	mF_Mpc_f_a: ARRAY[0..59047] OF LREAL := [-1.7756006070928429E-5, -1.955926027849794E-5, -2.1265642444599059E-5, -2.2878087249309936E-5, -2.4399475238503513E-5, -2.5832632877734329E-5, -2.7180332648224444E-5, -2.8445293182983732E-5, -2.9630179441154765E-5, -3.0737602918726609E-5, -3.1770121893815045E-5, -3.2730241704758869E-5, -3.3620415059333691E-5, -3.4443042373434618E-5, -3.5200472137629193E-5, -3.5895001310030509E-5, -3.652887573398812E-5, -3.7104290579141277E-5, -3.7623390804425058E-5, -3.808827164166491E-5, -3.8500979098439383E-5, -3.886351047893401E-5, -3.9177814921551905E-5, -3.9445793952087749E-5, -3.966930205131298E-5, -3.98501472358593E-5, -3.9990091651326829E-5, -4.0090852176581095E-5, -4.0154101038240283E-5, -4.0181466434390562E-5, -4.017453316660271E-5, -4.013484327935801E-5, -4.0063896706025282E-5, -3.9963151920563813E-5, -3.9834026594159355E-5, -3.9677898256031791E-5, -3.9496104957683613E-5, -3.9289945939888413E-5, -3.9060682301747689E-5, -3.8809537671172525E-5, -3.8537698876174604E-5, -3.8246316616377579E-5, -3.793650613418646E-5, -3.7609347885077623E-5, -3.7265888206497395E-5, -3.6907139984880808E-5, -3.6534083320325723E-5, -3.6147666188480321E-5, -3.5748805099224027E-5, -3.5338385751743129E-5, -3.4917263685623729E-5, -3.44862649276042E-5, -3.40461866336495E-5, -3.3597797726028135E-5, -3.3141839525091535E-5, -3.2679026375472935E-5, -3.221004626644033E-5, -3.1735561446154833E-5, -3.12562090296018E-5, -3.0772601599977736E-5, -3.0285327803331116E-5, -2.9794952936269942E-5, -2.9302019526562752E-5, -2.8807047906473585E-5, -2.8310536778684464E-5, -2.7812963774671571E-5, -2.7314786005413577E-5, -2.6816440604322343E-5, -2.6318345262297408E-5, -2.5820898754816765E-5, -2.5324481460986734E-5, -2.4829455874483883E-5, -2.4336167106331684E-5, -2.3844943379463754E-5, -2.3356096515034559E-5, -2.2869922410446928E-5, -2.2386701509073987E-5, -2.190669926166088E-5, -2.1430166579399207E-5, -2.0957340278674263E-5, -2.0488443517492027E-5, -2.0023686223599328E-5, -1.9563265514316956E-5, -1.910736610811127E-5, -1.8656160727935741E-5, -1.8209810496378919E-5, -1.776846532266075E-5, -1.7332264281523728E-5, -1.6901335984070202E-5, -1.6475798940601218E-5, -1.6055761915516631E-5, -1.5641324274339943E-5, -1.5232576322934952E-5, -1.4829599638984815E-5, -1.4432467395807249E-5, -1.4041244678582621E-5, -1.3655988793074526E-5, -1.3276749566924981E-5, -1.29035696436089E-5, -1.2536484769134677E-5, -1.217552407157984E-5, -1.1820710333552607E-5, -1.1472060257671982E-5, -1.1129584725160594E-5, -1.0793289047645905E-5, -1.0463173212266783E-5, -1.0139232120183559E-5, -9.8214558185907186E-6, -9.5098297263323067E-6, -9.20433485322091E-6, -8.9049480131616991E-6, -8.6116420311836354E-6, -8.324385944480339E-6, -8.04314519756346E-6, -7.7678818316316609E-6, -7.4985546682584246E-6, -7.2351194875019937E-6, -6.9775292005406626E-6, -6.7257340169365817E-6, -6.4796816066309883E-6, 1.7756006070928429E-5, 1.955926027849794E-5, 2.1265642444599059E-5, 2.2878087249309936E-5, 2.4399475238503513E-5, 2.5832632877734329E-5, 2.7180332648224444E-5, 2.8445293182983732E-5, 2.9630179441154765E-5, 3.0737602918726609E-5, 3.1770121893815045E-5, 3.2730241704758869E-5, 3.3620415059333691E-5, 3.4443042373434618E-5, 3.5200472137629193E-5, 3.5895001310030509E-5, 3.652887573398812E-5, 3.7104290579141277E-5, 3.7623390804425058E-5, 3.808827164166491E-5, 3.8500979098439383E-5, 3.886351047893401E-5, 3.9177814921551905E-5, 3.9445793952087749E-5, 3.966930205131298E-5, 3.98501472358593E-5, 3.9990091651326829E-5, 4.0090852176581095E-5, 4.0154101038240283E-5, 4.0181466434390562E-5, 4.017453316660271E-5, 4.013484327935801E-5, 4.0063896706025282E-5, 3.9963151920563813E-5, 3.9834026594159355E-5, 3.9677898256031791E-5, 3.9496104957683613E-5, 3.9289945939888413E-5, 3.9060682301747689E-5, 3.8809537671172525E-5, 3.8537698876174604E-5, 3.8246316616377579E-5, 3.793650613418646E-5, 3.7609347885077623E-5, 3.7265888206497395E-5, 3.6907139984880808E-5, 3.6534083320325723E-5, 3.6147666188480321E-5, 3.5748805099224027E-5, 3.5338385751743129E-5, 3.4917263685623729E-5, 3.44862649276042E-5, 3.40461866336495E-5, 3.3597797726028135E-5, 3.3141839525091535E-5, 3.2679026375472935E-5, 3.221004626644033E-5, 3.1735561446154833E-5, 3.12562090296018E-5, 3.0772601599977736E-5, 3.0285327803331116E-5, 2.9794952936269942E-5, 2.9302019526562752E-5, 2.8807047906473585E-5, 2.8310536778684464E-5, 2.7812963774671571E-5, 2.7314786005413577E-5, 2.6816440604322343E-5, 2.6318345262297408E-5, 2.5820898754816765E-5, 2.5324481460986734E-5, 2.4829455874483883E-5, 2.4336167106331684E-5, 2.3844943379463754E-5, 2.3356096515034559E-5, 2.2869922410446928E-5, 2.2386701509073987E-5, 2.190669926166088E-5, 2.1430166579399207E-5, 2.0957340278674263E-5, 2.0488443517492027E-5, 2.0023686223599328E-5, 1.9563265514316956E-5, 1.910736610811127E-5, 1.8656160727935741E-5, 1.8209810496378919E-5, 1.776846532266075E-5, 1.7332264281523728E-5, 1.6901335984070202E-5, 1.6475798940601218E-5, 1.6055761915516631E-5, 1.5641324274339943E-5, 1.5232576322934952E-5, 1.4829599638984815E-5, 1.4432467395807249E-5, 1.4041244678582621E-5, 1.3655988793074526E-5, 1.3276749566924981E-5, 1.29035696436089E-5, 1.2536484769134677E-5, 1.217552407157984E-5, 1.1820710333552607E-5, 1.1472060257671982E-5, 1.1129584725160594E-5, 1.0793289047645905E-5, 1.0463173212266783E-5, 1.0139232120183559E-5, 9.8214558185907186E-6, 9.5098297263323067E-6, 9.20433485322091E-6, 8.9049480131616991E-6, 8.6116420311836354E-6, 8.324385944480339E-6, 8.04314519756346E-6, 7.7678818316316609E-6, 7.4985546682584246E-6, 7.2351194875019937E-6, 6.9775292005406626E-6, 6.7257340169365817E-6, 6.4796816066309883E-6, 0.0, 0.0, 0.0, 0.0, -0.0, -0.0, -0.0, -0.0, -0.0, -0.0, -0.0, -0.0, -0.0, -0.0, -0.0, -0.0, -0.0, -0.0, -0.0, -0.0, -0.0, -0.0, -0.0, -0.0, -0.0, -0.0, -0.0, -0.0, -0.0, -0.0, -0.0, -0.0, -0.0, -0.0, -0.0, -0.0, -0.0, -0.0, -0.0, -0.0, -0.0, -0.0, -0.0, -0.0, -0.0, -0.0, -0.0, -0.0, -0.0, -0.0, -0.0, -0.0, -0.0, -0.0, -0.0, -0.0, -0.0, -0.0, -0.0, -0.0, -0.0, -0.0, -0.0, -0.0, -0.0, -0.0, -0.0, -0.0, -0.0, -0.0, -0.0, -0.0, -0.0, -0.0, -0.0, -0.0, -0.0, -0.0, -0.0, -0.0, -0.0, -0.0, -0.0, -0.0, -0.0, -0.0, -0.0, -0.0, -0.0, -0.0, -0.0, -0.0, -0.0, -0.0, -0.0, -0.0, -0.0, -0.0, -0.0, -0.0, -0.0, -0.0, -0.0, -0.0, -0.0, -0.0, -0.0, -0.0, -0.0, -0.0, -0.0, -0.0, -0.0, -0.0, -0.0, -0.0, -0.0, -0.0, -0.0, -0.0, -0.0, -0.0, -0.0, -0.0, 0.0, 0.0, 0.0, 0.0, 0.0, 0.0, 0.0, 0.0, 0.0, 0.0, 0.0, 0.0, 0.0, 0.0, 0.0, 0.0, 0.0, 0.0, 0.0, 0.0, 0.0, 0.0, 0.0, 0.0, 0.0, 0.0, 0.0, 0.0, 0.0, 0.0, 0.0, 0.0, 0.0, 0.0, 0.0, 0.0, 0.0, 0.0, 0.0, 0.0, 0.0, 0.0, 0.0, 0.0, 0.0, 0.0, 0.0, 0.0, 0.0, 0.0, 0.0, 0.0, 0.0, 0.0, 0.0, 0.0, 0.0, 0.0, 0.0, 0.0, 0.0, 0.0, 0.0, 0.0, 0.0, 0.0, 0.0, 0.0, 0.0, 0.0, 0.0, 0.0, 0.0, 0.0, 0.0, 0.0, 0.0, 0.0, 0.0, 0.0, 0.0, 0.0, 0.0, 0.0, 0.0, 0.0, 0.0, 0.0, 0.0, 0.0, 0.0, 0.0, 0.0, 0.0, 0.0, 0.0, 0.0, 0.0, 0.0, 0.0, 0.0, 0.0, 0.0, 0.0, 0.0, 0.0, 0.0, 0.0, 0.0, 0.0, 0.0, 0.0, 0.0, 0.0, 0.0, 0.0, 0.0, 0.0, 0.0, 0.0, 0.0, 0.0, 0.0, 0.0, -0.0, -1.7756006070928429E-5, -1.955926027849794E-5, -2.1265642444599059E-5, -2.2878087249309936E-5, -2.4399475238503513E-5, -2.5832632877734329E-5, -2.7180332648224444E-5, -2.8445293182983732E-5, -2.9630179441154765E-5, -3.0737602918726609E-5, -3.1770121893815045E-5, -3.2730241704758869E-5, -3.3620415059333691E-5, -3.4443042373434618E-5, -3.5200472137629193E-5, -3.5895001310030509E-5, -3.652887573398812E-5, -3.7104290579141277E-5, -3.7623390804425058E-5, -3.808827164166491E-5, -3.8500979098439383E-5, -3.886351047893401E-5, -3.9177814921551905E-5, -3.9445793952087749E-5, -3.966930205131298E-5, -3.98501472358593E-5, -3.9990091651326829E-5, -4.0090852176581095E-5, -4.0154101038240283E-5, -4.0181466434390562E-5, -4.017453316660271E-5, -4.013484327935801E-5, -4.0063896706025282E-5, -3.9963151920563813E-5, -3.9834026594159355E-5, -3.9677898256031791E-5, -3.9496104957683613E-5, -3.9289945939888413E-5, -3.9060682301747689E-5, -3.8809537671172525E-5, -3.8537698876174604E-5, -3.8246316616377579E-5, -3.793650613418646E-5, -3.7609347885077623E-5, -3.7265888206497395E-5, -3.6907139984880808E-5, -3.6534083320325723E-5, -3.6147666188480321E-5, -3.5748805099224027E-5, -3.5338385751743129E-5, -3.4917263685623729E-5, -3.44862649276042E-5, -3.40461866336495E-5, -3.3597797726028135E-5, -3.3141839525091535E-5, -3.2679026375472935E-5, -3.221004626644033E-5, -3.1735561446154833E-5, -3.12562090296018E-5, -3.0772601599977736E-5, -3.0285327803331116E-5, -2.9794952936269942E-5, -2.9302019526562752E-5, -2.8807047906473585E-5, -2.8310536778684464E-5, -2.7812963774671571E-5, -2.7314786005413577E-5, -2.6816440604322343E-5, -2.6318345262297408E-5, -2.5820898754816765E-5, -2.5324481460986734E-5, -2.4829455874483883E-5, -2.4336167106331684E-5, -2.3844943379463754E-5, -2.3356096515034559E-5, -2.2869922410446928E-5, -2.2386701509073987E-5, -2.190669926166088E-5, -2.1430166579399207E-5, -2.0957340278674263E-5, -2.0488443517492027E-5, -2.0023686223599328E-5, -1.9563265514316956E-5, -1.910736610811127E-5, -1.8656160727935741E-5, -1.8209810496378919E-5, -1.776846532266075E-5, -1.7332264281523728E-5, -1.6901335984070202E-5, -1.6475798940601218E-5, -1.6055761915516631E-5, -1.5641324274339943E-5, -1.5232576322934952E-5, -1.4829599638984815E-5, -1.4432467395807249E-5, -1.4041244678582621E-5, -1.3655988793074526E-5, -1.3276749566924981E-5, -1.29035696436089E-5, -1.2536484769134677E-5, -1.217552407157984E-5, -1.1820710333552607E-5, -1.1472060257671982E-5, -1.1129584725160594E-5, -1.0793289047645905E-5, -1.0463173212266783E-5, -1.0139232120183559E-5, -9.8214558185907186E-6, -9.5098297263323067E-6, -9.20433485322091E-6, -8.9049480131616991E-6, -8.6116420311836354E-6, -8.324385944480339E-6, -8.04314519756346E-6, -7.7678818316316609E-6, -7.4985546682584246E-6, -7.2351194875019937E-6, -6.9775292005406626E-6, -6.7257340169365817E-6, 0.0, 1.7756006070928429E-5, 1.955926027849794E-5, 2.1265642444599059E-5, 2.2878087249309936E-5, 2.4399475238503513E-5, 2.5832632877734329E-5, 2.7180332648224444E-5, 2.8445293182983732E-5, 2.9630179441154765E-5, 3.0737602918726609E-5, 3.1770121893815045E-5, 3.2730241704758869E-5, 3.3620415059333691E-5, 3.4443042373434618E-5, 3.5200472137629193E-5, 3.5895001310030509E-5, 3.652887573398812E-5, 3.7104290579141277E-5, 3.7623390804425058E-5, 3.808827164166491E-5, 3.8500979098439383E-5, 3.886351047893401E-5, 3.9177814921551905E-5, 3.9445793952087749E-5, 3.966930205131298E-5, 3.98501472358593E-5, 3.9990091651326829E-5, 4.0090852176581095E-5, 4.0154101038240283E-5, 4.0181466434390562E-5, 4.017453316660271E-5, 4.013484327935801E-5, 4.0063896706025282E-5, 3.9963151920563813E-5, 3.9834026594159355E-5, 3.9677898256031791E-5, 3.9496104957683613E-5, 3.9289945939888413E-5, 3.9060682301747689E-5, 3.8809537671172525E-5, 3.8537698876174604E-5, 3.8246316616377579E-5, 3.793650613418646E-5, 3.7609347885077623E-5, 3.7265888206497395E-5, 3.6907139984880808E-5, 3.6534083320325723E-5, 3.6147666188480321E-5, 3.5748805099224027E-5, 3.5338385751743129E-5, 3.4917263685623729E-5, 3.44862649276042E-5, 3.40461866336495E-5, 3.3597797726028135E-5, 3.3141839525091535E-5, 3.2679026375472935E-5, 3.221004626644033E-5, 3.1735561446154833E-5, 3.12562090296018E-5, 3.0772601599977736E-5, 3.0285327803331116E-5, 2.9794952936269942E-5, 2.9302019526562752E-5, 2.8807047906473585E-5, 2.8310536778684464E-5, 2.7812963774671571E-5, 2.7314786005413577E-5, 2.6816440604322343E-5, 2.6318345262297408E-5, 2.5820898754816765E-5, 2.5324481460986734E-5, 2.4829455874483883E-5, 2.4336167106331684E-5, 2.3844943379463754E-5, 2.3356096515034559E-5, 2.2869922410446928E-5, 2.2386701509073987E-5, 2.190669926166088E-5, 2.1430166579399207E-5, 2.0957340278674263E-5, 2.0488443517492027E-5, 2.0023686223599328E-5, 1.9563265514316956E-5, 1.910736610811127E-5, 1.8656160727935741E-5, 1.8209810496378919E-5, 1.776846532266075E-5, 1.7332264281523728E-5, 1.6901335984070202E-5, 1.6475798940601218E-5, 1.6055761915516631E-5, 1.5641324274339943E-5, 1.5232576322934952E-5, 1.4829599638984815E-5, 1.4432467395807249E-5, 1.4041244678582621E-5, 1.3655988793074526E-5, 1.3276749566924981E-5, 1.29035696436089E-5, 1.2536484769134677E-5, 1.217552407157984E-5, 1.1820710333552607E-5, 1.1472060257671982E-5, 1.1129584725160594E-5, 1.0793289047645905E-5, 1.0463173212266783E-5, 1.0139232120183559E-5, 9.8214558185907186E-6, 9.5098297263323067E-6, 9.20433485322091E-6, 8.9049480131616991E-6, 8.6116420311836354E-6, 8.324385944480339E-6, 8.04314519756346E-6, 7.7678818316316609E-6, 7.4985546682584246E-6, 7.2351194875019937E-6, 6.9775292005406626E-6, 6.7257340169365817E-6, 0.0, 0.0, 0.0, 0.0, -0.0, -0.0, -0.0, -0.0, -0.0, -0.0, -0.0, -0.0, -0.0, -0.0, -0.0, -0.0, -0.0, -0.0, -0.0, -0.0, -0.0, -0.0, -0.0, -0.0, -0.0, -0.0, -0.0, -0.0, -0.0, -0.0, -0.0, -0.0, -0.0, -0.0, -0.0, -0.0, -0.0, -0.0, -0.0, -0.0, -0.0, -0.0, -0.0, -0.0, -0.0, -0.0, -0.0, -0.0, -0.0, -0.0, -0.0, -0.0, -0.0, -0.0, -0.0, -0.0, -0.0, -0.0, -0.0, -0.0, -0.0, -0.0, -0.0, -0.0, -0.0, -0.0, -0.0, -0.0, -0.0, -0.0, -0.0, -0.0, -0.0, -0.0, -0.0, -0.0, -0.0, -0.0, -0.0, -0.0, -0.0, -0.0, -0.0, -0.0, -0.0, -0.0, -0.0, -0.0, -0.0, -0.0, -0.0, -0.0, -0.0, -0.0, -0.0, -0.0, -0.0, -0.0, -0.0, -0.0, -0.0, -0.0, -0.0, -0.0, -0.0, -0.0, -0.0, -0.0, -0.0, -0.0, -0.0, -0.0, -0.0, -0.0, -0.0, -0.0, -0.0, -0.0, -0.0, -0.0, -0.0, -0.0, -0.0, -0.0, 0.0, 0.0, 0.0, 0.0, 0.0, 0.0, 0.0, 0.0, 0.0, 0.0, 0.0, 0.0, 0.0, 0.0, 0.0, 0.0, 0.0, 0.0, 0.0, 0.0, 0.0, 0.0, 0.0, 0.0, 0.0, 0.0, 0.0, 0.0, 0.0, 0.0, 0.0, 0.0, 0.0, 0.0, 0.0, 0.0, 0.0, 0.0, 0.0, 0.0, 0.0, 0.0, 0.0, 0.0, 0.0, 0.0, 0.0, 0.0, 0.0, 0.0, 0.0, 0.0, 0.0, 0.0, 0.0, 0.0, 0.0, 0.0, 0.0, 0.0, 0.0, 0.0, 0.0, 0.0, 0.0, 0.0, 0.0, 0.0, 0.0, 0.0, 0.0, 0.0, 0.0, 0.0, 0.0, 0.0, 0.0, 0.0, 0.0, 0.0, 0.0, 0.0, 0.0, 0.0, 0.0, 0.0, 0.0, 0.0, 0.0, 0.0, 0.0, 0.0, 0.0, 0.0, 0.0, 0.0, 0.0, 0.0, 0.0, 0.0, 0.0, 0.0, 0.0, 0.0, 0.0, 0.0, 0.0, 0.0, 0.0, 0.0, 0.0, 0.0, 0.0, 0.0, 0.0, 0.0, 0.0, 0.0, 0.0, 0.0, 0.0, 0.0, 0.0, 0.0, -0.0, -0.0, -1.7756006070928429E-5, -1.955926027849794E-5, -2.1265642444599059E-5, -2.2878087249309936E-5, -2.4399475238503513E-5, -2.5832632877734329E-5, -2.7180332648224444E-5, -2.8445293182983732E-5, -2.9630179441154765E-5, -3.0737602918726609E-5, -3.1770121893815045E-5, -3.2730241704758869E-5, -3.3620415059333691E-5, -3.4443042373434618E-5, -3.5200472137629193E-5, -3.5895001310030509E-5, -3.652887573398812E-5, -3.7104290579141277E-5, -3.7623390804425058E-5, -3.808827164166491E-5, -3.8500979098439383E-5, -3.886351047893401E-5, -3.9177814921551905E-5, -3.9445793952087749E-5, -3.966930205131298E-5, -3.98501472358593E-5, -3.9990091651326829E-5, -4.0090852176581095E-5, -4.0154101038240283E-5, -4.0181466434390562E-5, -4.017453316660271E-5, -4.013484327935801E-5, -4.0063896706025282E-5, -3.9963151920563813E-5, -3.9834026594159355E-5, -3.9677898256031791E-5, -3.9496104957683613E-5, -3.9289945939888413E-5, -3.9060682301747689E-5, -3.8809537671172525E-5, -3.8537698876174604E-5, -3.8246316616377579E-5, -3.793650613418646E-5, -3.7609347885077623E-5, -3.7265888206497395E-5, -3.6907139984880808E-5, -3.6534083320325723E-5, -3.6147666188480321E-5, -3.5748805099224027E-5, -3.5338385751743129E-5, -3.4917263685623729E-5, -3.44862649276042E-5, -3.40461866336495E-5, -3.3597797726028135E-5, -3.3141839525091535E-5, -3.2679026375472935E-5, -3.221004626644033E-5, -3.1735561446154833E-5, -3.12562090296018E-5, -3.0772601599977736E-5, -3.0285327803331116E-5, -2.9794952936269942E-5, -2.9302019526562752E-5, -2.8807047906473585E-5, -2.8310536778684464E-5, -2.7812963774671571E-5, -2.7314786005413577E-5, -2.6816440604322343E-5, -2.6318345262297408E-5, -2.5820898754816765E-5, -2.5324481460986734E-5, -2.4829455874483883E-5, -2.4336167106331684E-5, -2.3844943379463754E-5, -2.3356096515034559E-5, -2.2869922410446928E-5, -2.2386701509073987E-5, -2.190669926166088E-5, -2.1430166579399207E-5, -2.0957340278674263E-5, -2.0488443517492027E-5, -2.0023686223599328E-5, -1.9563265514316956E-5, -1.910736610811127E-5, -1.8656160727935741E-5, -1.8209810496378919E-5, -1.776846532266075E-5, -1.7332264281523728E-5, -1.6901335984070202E-5, -1.6475798940601218E-5, -1.6055761915516631E-5, -1.5641324274339943E-5, -1.5232576322934952E-5, -1.4829599638984815E-5, -1.4432467395807249E-5, -1.4041244678582621E-5, -1.3655988793074526E-5, -1.3276749566924981E-5, -1.29035696436089E-5, -1.2536484769134677E-5, -1.217552407157984E-5, -1.1820710333552607E-5, -1.1472060257671982E-5, -1.1129584725160594E-5, -1.0793289047645905E-5, -1.0463173212266783E-5, -1.0139232120183559E-5, -9.8214558185907186E-6, -9.5098297263323067E-6, -9.20433485322091E-6, -8.9049480131616991E-6, -8.6116420311836354E-6, -8.324385944480339E-6, -8.04314519756346E-6, -7.7678818316316609E-6, -7.4985546682584246E-6, -7.2351194875019937E-6, -6.9775292005406626E-6, 0.0, 0.0, 1.7756006070928429E-5, 1.955926027849794E-5, 2.1265642444599059E-5, 2.2878087249309936E-5, 2.4399475238503513E-5, 2.5832632877734329E-5, 2.7180332648224444E-5, 2.8445293182983732E-5, 2.9630179441154765E-5, 3.0737602918726609E-5, 3.1770121893815045E-5, 3.2730241704758869E-5, 3.3620415059333691E-5, 3.4443042373434618E-5, 3.5200472137629193E-5, 3.5895001310030509E-5, 3.652887573398812E-5, 3.7104290579141277E-5, 3.7623390804425058E-5, 3.808827164166491E-5, 3.8500979098439383E-5, 3.886351047893401E-5, 3.9177814921551905E-5, 3.9445793952087749E-5, 3.966930205131298E-5, 3.98501472358593E-5, 3.9990091651326829E-5, 4.0090852176581095E-5, 4.0154101038240283E-5, 4.0181466434390562E-5, 4.017453316660271E-5, 4.013484327935801E-5, 4.0063896706025282E-5, 3.9963151920563813E-5, 3.9834026594159355E-5, 3.9677898256031791E-5, 3.9496104957683613E-5, 3.9289945939888413E-5, 3.9060682301747689E-5, 3.8809537671172525E-5, 3.8537698876174604E-5, 3.8246316616377579E-5, 3.793650613418646E-5, 3.7609347885077623E-5, 3.7265888206497395E-5, 3.6907139984880808E-5, 3.6534083320325723E-5, 3.6147666188480321E-5, 3.5748805099224027E-5, 3.5338385751743129E-5, 3.4917263685623729E-5, 3.44862649276042E-5, 3.40461866336495E-5, 3.3597797726028135E-5, 3.3141839525091535E-5, 3.2679026375472935E-5, 3.221004626644033E-5, 3.1735561446154833E-5, 3.12562090296018E-5, 3.0772601599977736E-5, 3.0285327803331116E-5, 2.9794952936269942E-5, 2.9302019526562752E-5, 2.8807047906473585E-5, 2.8310536778684464E-5, 2.7812963774671571E-5, 2.7314786005413577E-5, 2.6816440604322343E-5, 2.6318345262297408E-5, 2.5820898754816765E-5, 2.5324481460986734E-5, 2.4829455874483883E-5, 2.4336167106331684E-5, 2.3844943379463754E-5, 2.3356096515034559E-5, 2.2869922410446928E-5, 2.2386701509073987E-5, 2.190669926166088E-5, 2.1430166579399207E-5, 2.0957340278674263E-5, 2.0488443517492027E-5, 2.0023686223599328E-5, 1.9563265514316956E-5, 1.910736610811127E-5, 1.8656160727935741E-5, 1.8209810496378919E-5, 1.776846532266075E-5, 1.7332264281523728E-5, 1.6901335984070202E-5, 1.6475798940601218E-5, 1.6055761915516631E-5, 1.5641324274339943E-5, 1.5232576322934952E-5, 1.4829599638984815E-5, 1.4432467395807249E-5, 1.4041244678582621E-5, 1.3655988793074526E-5, 1.3276749566924981E-5, 1.29035696436089E-5, 1.2536484769134677E-5, 1.217552407157984E-5, 1.1820710333552607E-5, 1.1472060257671982E-5, 1.1129584725160594E-5, 1.0793289047645905E-5, 1.0463173212266783E-5, 1.0139232120183559E-5, 9.8214558185907186E-6, 9.5098297263323067E-6, 9.20433485322091E-6, 8.9049480131616991E-6, 8.6116420311836354E-6, 8.324385944480339E-6, 8.04314519756346E-6, 7.7678818316316609E-6, 7.4985546682584246E-6, 7.2351194875019937E-6, 6.9775292005406626E-6, 0.0, 0.0, 0.0, 0.0, -0.0, -0.0, -0.0, -0.0, -0.0, -0.0, -0.0, -0.0, -0.0, -0.0, -0.0, -0.0, -0.0, -0.0, -0.0, -0.0, -0.0, -0.0, -0.0, -0.0, -0.0, -0.0, -0.0, -0.0, -0.0, -0.0, -0.0, -0.0, -0.0, -0.0, -0.0, -0.0, -0.0, -0.0, -0.0, -0.0, -0.0, -0.0, -0.0, -0.0, -0.0, -0.0, -0.0, -0.0, -0.0, -0.0, -0.0, -0.0, -0.0, -0.0, -0.0, -0.0, -0.0, -0.0, -0.0, -0.0, -0.0, -0.0, -0.0, -0.0, -0.0, -0.0, -0.0, -0.0, -0.0, -0.0, -0.0, -0.0, -0.0, -0.0, -0.0, -0.0, -0.0, -0.0, -0.0, -0.0, -0.0, -0.0, -0.0, -0.0, -0.0, -0.0, -0.0, -0.0, -0.0, -0.0, -0.0, -0.0, -0.0, -0.0, -0.0, -0.0, -0.0, -0.0, -0.0, -0.0, -0.0, -0.0, -0.0, -0.0, -0.0, -0.0, -0.0, -0.0, -0.0, -0.0, -0.0, -0.0, -0.0, -0.0, -0.0, -0.0, -0.0, -0.0, -0.0, -0.0, -0.0, -0.0, -0.0, -0.0, 0.0, 0.0, 0.0, 0.0, 0.0, 0.0, 0.0, 0.0, 0.0, 0.0, 0.0, 0.0, 0.0, 0.0, 0.0, 0.0, 0.0, 0.0, 0.0, 0.0, 0.0, 0.0, 0.0, 0.0, 0.0, 0.0, 0.0, 0.0, 0.0, 0.0, 0.0, 0.0, 0.0, 0.0, 0.0, 0.0, 0.0, 0.0, 0.0, 0.0, 0.0, 0.0, 0.0, 0.0, 0.0, 0.0, 0.0, 0.0, 0.0, 0.0, 0.0, 0.0, 0.0, 0.0, 0.0, 0.0, 0.0, 0.0, 0.0, 0.0, 0.0, 0.0, 0.0, 0.0, 0.0, 0.0, 0.0, 0.0, 0.0, 0.0, 0.0, 0.0, 0.0, 0.0, 0.0, 0.0, 0.0, 0.0, 0.0, 0.0, 0.0, 0.0, 0.0, 0.0, 0.0, 0.0, 0.0, 0.0, 0.0, 0.0, 0.0, 0.0, 0.0, 0.0, 0.0, 0.0, 0.0, 0.0, 0.0, 0.0, 0.0, 0.0, 0.0, 0.0, 0.0, 0.0, 0.0, 0.0, 0.0, 0.0, 0.0, 0.0, 0.0, 0.0, 0.0, 0.0, 0.0, 0.0, 0.0, 0.0, 0.0, 0.0, 0.0, 0.0, -0.0, -0.0, -0.0, -1.7756006070928429E-5, -1.955926027849794E-5, -2.1265642444599059E-5, -2.2878087249309936E-5, -2.4399475238503513E-5, -2.5832632877734329E-5, -2.7180332648224444E-5, -2.8445293182983732E-5, -2.9630179441154765E-5, -3.0737602918726609E-5, -3.1770121893815045E-5, -3.2730241704758869E-5, -3.3620415059333691E-5, -3.4443042373434618E-5, -3.5200472137629193E-5, -3.5895001310030509E-5, -3.652887573398812E-5, -3.7104290579141277E-5, -3.7623390804425058E-5, -3.808827164166491E-5, -3.8500979098439383E-5, -3.886351047893401E-5, -3.9177814921551905E-5, -3.9445793952087749E-5, -3.966930205131298E-5, -3.98501472358593E-5, -3.9990091651326829E-5, -4.0090852176581095E-5, -4.0154101038240283E-5, -4.0181466434390562E-5, -4.017453316660271E-5, -4.013484327935801E-5, -4.0063896706025282E-5, -3.9963151920563813E-5, -3.9834026594159355E-5, -3.9677898256031791E-5, -3.9496104957683613E-5, -3.9289945939888413E-5, -3.9060682301747689E-5, -3.8809537671172525E-5, -3.8537698876174604E-5, -3.8246316616377579E-5, -3.793650613418646E-5, -3.7609347885077623E-5, -3.7265888206497395E-5, -3.6907139984880808E-5, -3.6534083320325723E-5, -3.6147666188480321E-5, -3.5748805099224027E-5, -3.5338385751743129E-5, -3.4917263685623729E-5, -3.44862649276042E-5, -3.40461866336495E-5, -3.3597797726028135E-5, -3.3141839525091535E-5, -3.2679026375472935E-5, -3.221004626644033E-5, -3.1735561446154833E-5, -3.12562090296018E-5, -3.0772601599977736E-5, -3.0285327803331116E-5, -2.9794952936269942E-5, -2.9302019526562752E-5, -2.8807047906473585E-5, -2.8310536778684464E-5, -2.7812963774671571E-5, -2.7314786005413577E-5, -2.6816440604322343E-5, -2.6318345262297408E-5, -2.5820898754816765E-5, -2.5324481460986734E-5, -2.4829455874483883E-5, -2.4336167106331684E-5, -2.3844943379463754E-5, -2.3356096515034559E-5, -2.2869922410446928E-5, -2.2386701509073987E-5, -2.190669926166088E-5, -2.1430166579399207E-5, -2.0957340278674263E-5, -2.0488443517492027E-5, -2.0023686223599328E-5, -1.9563265514316956E-5, -1.910736610811127E-5, -1.8656160727935741E-5, -1.8209810496378919E-5, -1.776846532266075E-5, -1.7332264281523728E-5, -1.6901335984070202E-5, -1.6475798940601218E-5, -1.6055761915516631E-5, -1.5641324274339943E-5, -1.5232576322934952E-5, -1.4829599638984815E-5, -1.4432467395807249E-5, -1.4041244678582621E-5, -1.3655988793074526E-5, -1.3276749566924981E-5, -1.29035696436089E-5, -1.2536484769134677E-5, -1.217552407157984E-5, -1.1820710333552607E-5, -1.1472060257671982E-5, -1.1129584725160594E-5, -1.0793289047645905E-5, -1.0463173212266783E-5, -1.0139232120183559E-5, -9.8214558185907186E-6, -9.5098297263323067E-6, -9.20433485322091E-6, -8.9049480131616991E-6, -8.6116420311836354E-6, -8.324385944480339E-6, -8.04314519756346E-6, -7.7678818316316609E-6, -7.4985546682584246E-6, -7.2351194875019937E-6, 0.0, 0.0, 0.0, 1.7756006070928429E-5, 1.955926027849794E-5, 2.1265642444599059E-5, 2.2878087249309936E-5, 2.4399475238503513E-5, 2.5832632877734329E-5, 2.7180332648224444E-5, 2.8445293182983732E-5, 2.9630179441154765E-5, 3.0737602918726609E-5, 3.1770121893815045E-5, 3.2730241704758869E-5, 3.3620415059333691E-5, 3.4443042373434618E-5, 3.5200472137629193E-5, 3.5895001310030509E-5, 3.652887573398812E-5, 3.7104290579141277E-5, 3.7623390804425058E-5, 3.808827164166491E-5, 3.8500979098439383E-5, 3.886351047893401E-5, 3.9177814921551905E-5, 3.9445793952087749E-5, 3.966930205131298E-5, 3.98501472358593E-5, 3.9990091651326829E-5, 4.0090852176581095E-5, 4.0154101038240283E-5, 4.0181466434390562E-5, 4.017453316660271E-5, 4.013484327935801E-5, 4.0063896706025282E-5, 3.9963151920563813E-5, 3.9834026594159355E-5, 3.9677898256031791E-5, 3.9496104957683613E-5, 3.9289945939888413E-5, 3.9060682301747689E-5, 3.8809537671172525E-5, 3.8537698876174604E-5, 3.8246316616377579E-5, 3.793650613418646E-5, 3.7609347885077623E-5, 3.7265888206497395E-5, 3.6907139984880808E-5, 3.6534083320325723E-5, 3.6147666188480321E-5, 3.5748805099224027E-5, 3.5338385751743129E-5, 3.4917263685623729E-5, 3.44862649276042E-5, 3.40461866336495E-5, 3.3597797726028135E-5, 3.3141839525091535E-5, 3.2679026375472935E-5, 3.221004626644033E-5, 3.1735561446154833E-5, 3.12562090296018E-5, 3.0772601599977736E-5, 3.0285327803331116E-5, 2.9794952936269942E-5, 2.9302019526562752E-5, 2.8807047906473585E-5, 2.8310536778684464E-5, 2.7812963774671571E-5, 2.7314786005413577E-5, 2.6816440604322343E-5, 2.6318345262297408E-5, 2.5820898754816765E-5, 2.5324481460986734E-5, 2.4829455874483883E-5, 2.4336167106331684E-5, 2.3844943379463754E-5, 2.3356096515034559E-5, 2.2869922410446928E-5, 2.2386701509073987E-5, 2.190669926166088E-5, 2.1430166579399207E-5, 2.0957340278674263E-5, 2.0488443517492027E-5, 2.0023686223599328E-5, 1.9563265514316956E-5, 1.910736610811127E-5, 1.8656160727935741E-5, 1.8209810496378919E-5, 1.776846532266075E-5, 1.7332264281523728E-5, 1.6901335984070202E-5, 1.6475798940601218E-5, 1.6055761915516631E-5, 1.5641324274339943E-5, 1.5232576322934952E-5, 1.4829599638984815E-5, 1.4432467395807249E-5, 1.4041244678582621E-5, 1.3655988793074526E-5, 1.3276749566924981E-5, 1.29035696436089E-5, 1.2536484769134677E-5, 1.217552407157984E-5, 1.1820710333552607E-5, 1.1472060257671982E-5, 1.1129584725160594E-5, 1.0793289047645905E-5, 1.0463173212266783E-5, 1.0139232120183559E-5, 9.8214558185907186E-6, 9.5098297263323067E-6, 9.20433485322091E-6, 8.9049480131616991E-6, 8.6116420311836354E-6, 8.324385944480339E-6, 8.04314519756346E-6, 7.7678818316316609E-6, 7.4985546682584246E-6, 7.2351194875019937E-6, 0.0, 0.0, 0.0, 0.0, -0.0, -0.0, -0.0, -0.0, -0.0, -0.0, -0.0, -0.0, -0.0, -0.0, -0.0, -0.0, -0.0, -0.0, -0.0, -0.0, -0.0, -0.0, -0.0, -0.0, -0.0, -0.0, -0.0, -0.0, -0.0, -0.0, -0.0, -0.0, -0.0, -0.0, -0.0, -0.0, -0.0, -0.0, -0.0, -0.0, -0.0, -0.0, -0.0, -0.0, -0.0, -0.0, -0.0, -0.0, -0.0, -0.0, -0.0, -0.0, -0.0, -0.0, -0.0, -0.0, -0.0, -0.0, -0.0, -0.0, -0.0, -0.0, -0.0, -0.0, -0.0, -0.0, -0.0, -0.0, -0.0, -0.0, -0.0, -0.0, -0.0, -0.0, -0.0, -0.0, -0.0, -0.0, -0.0, -0.0, -0.0, -0.0, -0.0, -0.0, -0.0, -0.0, -0.0, -0.0, -0.0, -0.0, -0.0, -0.0, -0.0, -0.0, -0.0, -0.0, -0.0, -0.0, -0.0, -0.0, -0.0, -0.0, -0.0, -0.0, -0.0, -0.0, -0.0, -0.0, -0.0, -0.0, -0.0, -0.0, -0.0, -0.0, -0.0, -0.0, -0.0, -0.0, -0.0, -0.0, -0.0, -0.0, -0.0, -0.0, 0.0, 0.0, 0.0, 0.0, 0.0, 0.0, 0.0, 0.0, 0.0, 0.0, 0.0, 0.0, 0.0, 0.0, 0.0, 0.0, 0.0, 0.0, 0.0, 0.0, 0.0, 0.0, 0.0, 0.0, 0.0, 0.0, 0.0, 0.0, 0.0, 0.0, 0.0, 0.0, 0.0, 0.0, 0.0, 0.0, 0.0, 0.0, 0.0, 0.0, 0.0, 0.0, 0.0, 0.0, 0.0, 0.0, 0.0, 0.0, 0.0, 0.0, 0.0, 0.0, 0.0, 0.0, 0.0, 0.0, 0.0, 0.0, 0.0, 0.0, 0.0, 0.0, 0.0, 0.0, 0.0, 0.0, 0.0, 0.0, 0.0, 0.0, 0.0, 0.0, 0.0, 0.0, 0.0, 0.0, 0.0, 0.0, 0.0, 0.0, 0.0, 0.0, 0.0, 0.0, 0.0, 0.0, 0.0, 0.0, 0.0, 0.0, 0.0, 0.0, 0.0, 0.0, 0.0, 0.0, 0.0, 0.0, 0.0, 0.0, 0.0, 0.0, 0.0, 0.0, 0.0, 0.0, 0.0, 0.0, 0.0, 0.0, 0.0, 0.0, 0.0, 0.0, 0.0, 0.0, 0.0, 0.0, 0.0, 0.0, 0.0, 0.0, 0.0, 0.0, -0.0, -0.0, -0.0, -0.0, -1.7756006070928429E-5, -1.955926027849794E-5, -2.1265642444599059E-5, -2.2878087249309936E-5, -2.4399475238503513E-5, -2.5832632877734329E-5, -2.7180332648224444E-5, -2.8445293182983732E-5, -2.9630179441154765E-5, -3.0737602918726609E-5, -3.1770121893815045E-5, -3.2730241704758869E-5, -3.3620415059333691E-5, -3.4443042373434618E-5, -3.5200472137629193E-5, -3.5895001310030509E-5, -3.652887573398812E-5, -3.7104290579141277E-5, -3.7623390804425058E-5, -3.808827164166491E-5, -3.8500979098439383E-5, -3.886351047893401E-5, -3.9177814921551905E-5, -3.9445793952087749E-5, -3.966930205131298E-5, -3.98501472358593E-5, -3.9990091651326829E-5, -4.0090852176581095E-5, -4.0154101038240283E-5, -4.0181466434390562E-5, -4.017453316660271E-5, -4.013484327935801E-5, -4.0063896706025282E-5, -3.9963151920563813E-5, -3.9834026594159355E-5, -3.9677898256031791E-5, -3.9496104957683613E-5, -3.9289945939888413E-5, -3.9060682301747689E-5, -3.8809537671172525E-5, -3.8537698876174604E-5, -3.8246316616377579E-5, -3.793650613418646E-5, -3.7609347885077623E-5, -3.7265888206497395E-5, -3.6907139984880808E-5, -3.6534083320325723E-5, -3.6147666188480321E-5, -3.5748805099224027E-5, -3.5338385751743129E-5, -3.4917263685623729E-5, -3.44862649276042E-5, -3.40461866336495E-5, -3.3597797726028135E-5, -3.3141839525091535E-5, -3.2679026375472935E-5, -3.221004626644033E-5, -3.1735561446154833E-5, -3.12562090296018E-5, -3.0772601599977736E-5, -3.0285327803331116E-5, -2.9794952936269942E-5, -2.9302019526562752E-5, -2.8807047906473585E-5, -2.8310536778684464E-5, -2.7812963774671571E-5, -2.7314786005413577E-5, -2.6816440604322343E-5, -2.6318345262297408E-5, -2.5820898754816765E-5, -2.5324481460986734E-5, -2.4829455874483883E-5, -2.4336167106331684E-5, -2.3844943379463754E-5, -2.3356096515034559E-5, -2.2869922410446928E-5, -2.2386701509073987E-5, -2.190669926166088E-5, -2.1430166579399207E-5, -2.0957340278674263E-5, -2.0488443517492027E-5, -2.0023686223599328E-5, -1.9563265514316956E-5, -1.910736610811127E-5, -1.8656160727935741E-5, -1.8209810496378919E-5, -1.776846532266075E-5, -1.7332264281523728E-5, -1.6901335984070202E-5, -1.6475798940601218E-5, -1.6055761915516631E-5, -1.5641324274339943E-5, -1.5232576322934952E-5, -1.4829599638984815E-5, -1.4432467395807249E-5, -1.4041244678582621E-5, -1.3655988793074526E-5, -1.3276749566924981E-5, -1.29035696436089E-5, -1.2536484769134677E-5, -1.217552407157984E-5, -1.1820710333552607E-5, -1.1472060257671982E-5, -1.1129584725160594E-5, -1.0793289047645905E-5, -1.0463173212266783E-5, -1.0139232120183559E-5, -9.8214558185907186E-6, -9.5098297263323067E-6, -9.20433485322091E-6, -8.9049480131616991E-6, -8.6116420311836354E-6, -8.324385944480339E-6, -8.04314519756346E-6, -7.7678818316316609E-6, -7.4985546682584246E-6, 0.0, 0.0, 0.0, 0.0, 1.7756006070928429E-5, 1.955926027849794E-5, 2.1265642444599059E-5, 2.2878087249309936E-5, 2.4399475238503513E-5, 2.5832632877734329E-5, 2.7180332648224444E-5, 2.8445293182983732E-5, 2.9630179441154765E-5, 3.0737602918726609E-5, 3.1770121893815045E-5, 3.2730241704758869E-5, 3.3620415059333691E-5, 3.4443042373434618E-5, 3.5200472137629193E-5, 3.5895001310030509E-5, 3.652887573398812E-5, 3.7104290579141277E-5, 3.7623390804425058E-5, 3.808827164166491E-5, 3.8500979098439383E-5, 3.886351047893401E-5, 3.9177814921551905E-5, 3.9445793952087749E-5, 3.966930205131298E-5, 3.98501472358593E-5, 3.9990091651326829E-5, 4.0090852176581095E-5, 4.0154101038240283E-5, 4.0181466434390562E-5, 4.017453316660271E-5, 4.013484327935801E-5, 4.0063896706025282E-5, 3.9963151920563813E-5, 3.9834026594159355E-5, 3.9677898256031791E-5, 3.9496104957683613E-5, 3.9289945939888413E-5, 3.9060682301747689E-5, 3.8809537671172525E-5, 3.8537698876174604E-5, 3.8246316616377579E-5, 3.793650613418646E-5, 3.7609347885077623E-5, 3.7265888206497395E-5, 3.6907139984880808E-5, 3.6534083320325723E-5, 3.6147666188480321E-5, 3.5748805099224027E-5, 3.5338385751743129E-5, 3.4917263685623729E-5, 3.44862649276042E-5, 3.40461866336495E-5, 3.3597797726028135E-5, 3.3141839525091535E-5, 3.2679026375472935E-5, 3.221004626644033E-5, 3.1735561446154833E-5, 3.12562090296018E-5, 3.0772601599977736E-5, 3.0285327803331116E-5, 2.9794952936269942E-5, 2.9302019526562752E-5, 2.8807047906473585E-5, 2.8310536778684464E-5, 2.7812963774671571E-5, 2.7314786005413577E-5, 2.6816440604322343E-5, 2.6318345262297408E-5, 2.5820898754816765E-5, 2.5324481460986734E-5, 2.4829455874483883E-5, 2.4336167106331684E-5, 2.3844943379463754E-5, 2.3356096515034559E-5, 2.2869922410446928E-5, 2.2386701509073987E-5, 2.190669926166088E-5, 2.1430166579399207E-5, 2.0957340278674263E-5, 2.0488443517492027E-5, 2.0023686223599328E-5, 1.9563265514316956E-5, 1.910736610811127E-5, 1.8656160727935741E-5, 1.8209810496378919E-5, 1.776846532266075E-5, 1.7332264281523728E-5, 1.6901335984070202E-5, 1.6475798940601218E-5, 1.6055761915516631E-5, 1.5641324274339943E-5, 1.5232576322934952E-5, 1.4829599638984815E-5, 1.4432467395807249E-5, 1.4041244678582621E-5, 1.3655988793074526E-5, 1.3276749566924981E-5, 1.29035696436089E-5, 1.2536484769134677E-5, 1.217552407157984E-5, 1.1820710333552607E-5, 1.1472060257671982E-5, 1.1129584725160594E-5, 1.0793289047645905E-5, 1.0463173212266783E-5, 1.0139232120183559E-5, 9.8214558185907186E-6, 9.5098297263323067E-6, 9.20433485322091E-6, 8.9049480131616991E-6, 8.6116420311836354E-6, 8.324385944480339E-6, 8.04314519756346E-6, 7.7678818316316609E-6, 7.4985546682584246E-6, 0.0, 0.0, 0.0, 0.0, -0.0, -0.0, -0.0, -0.0, -0.0, -0.0, -0.0, -0.0, -0.0, -0.0, -0.0, -0.0, -0.0, -0.0, -0.0, -0.0, -0.0, -0.0, -0.0, -0.0, -0.0, -0.0, -0.0, -0.0, -0.0, -0.0, -0.0, -0.0, -0.0, -0.0, -0.0, -0.0, -0.0, -0.0, -0.0, -0.0, -0.0, -0.0, -0.0, -0.0, -0.0, -0.0, -0.0, -0.0, -0.0, -0.0, -0.0, -0.0, -0.0, -0.0, -0.0, -0.0, -0.0, -0.0, -0.0, -0.0, -0.0, -0.0, -0.0, -0.0, -0.0, -0.0, -0.0, -0.0, -0.0, -0.0, -0.0, -0.0, -0.0, -0.0, -0.0, -0.0, -0.0, -0.0, -0.0, -0.0, -0.0, -0.0, -0.0, -0.0, -0.0, -0.0, -0.0, -0.0, -0.0, -0.0, -0.0, -0.0, -0.0, -0.0, -0.0, -0.0, -0.0, -0.0, -0.0, -0.0, -0.0, -0.0, -0.0, -0.0, -0.0, -0.0, -0.0, -0.0, -0.0, -0.0, -0.0, -0.0, -0.0, -0.0, -0.0, -0.0, -0.0, -0.0, -0.0, -0.0, -0.0, -0.0, -0.0, -0.0, 0.0, 0.0, 0.0, 0.0, 0.0, 0.0, 0.0, 0.0, 0.0, 0.0, 0.0, 0.0, 0.0, 0.0, 0.0, 0.0, 0.0, 0.0, 0.0, 0.0, 0.0, 0.0, 0.0, 0.0, 0.0, 0.0, 0.0, 0.0, 0.0, 0.0, 0.0, 0.0, 0.0, 0.0, 0.0, 0.0, 0.0, 0.0, 0.0, 0.0, 0.0, 0.0, 0.0, 0.0, 0.0, 0.0, 0.0, 0.0, 0.0, 0.0, 0.0, 0.0, 0.0, 0.0, 0.0, 0.0, 0.0, 0.0, 0.0, 0.0, 0.0, 0.0, 0.0, 0.0, 0.0, 0.0, 0.0, 0.0, 0.0, 0.0, 0.0, 0.0, 0.0, 0.0, 0.0, 0.0, 0.0, 0.0, 0.0, 0.0, 0.0, 0.0, 0.0, 0.0, 0.0, 0.0, 0.0, 0.0, 0.0, 0.0, 0.0, 0.0, 0.0, 0.0, 0.0, 0.0, 0.0, 0.0, 0.0, 0.0, 0.0, 0.0, 0.0, 0.0, 0.0, 0.0, 0.0, 0.0, 0.0, 0.0, 0.0, 0.0, 0.0, 0.0, 0.0, 0.0, 0.0, 0.0, 0.0, 0.0, 0.0, 0.0, 0.0, 0.0, -0.0, -0.0, -0.0, -0.0, -0.0, -1.7756006070928429E-5, -1.955926027849794E-5, -2.1265642444599059E-5, -2.2878087249309936E-5, -2.4399475238503513E-5, -2.5832632877734329E-5, -2.7180332648224444E-5, -2.8445293182983732E-5, -2.9630179441154765E-5, -3.0737602918726609E-5, -3.1770121893815045E-5, -3.2730241704758869E-5, -3.3620415059333691E-5, -3.4443042373434618E-5, -3.5200472137629193E-5, -3.5895001310030509E-5, -3.652887573398812E-5, -3.7104290579141277E-5, -3.7623390804425058E-5, -3.808827164166491E-5, -3.8500979098439383E-5, -3.886351047893401E-5, -3.9177814921551905E-5, -3.9445793952087749E-5, -3.966930205131298E-5, -3.98501472358593E-5, -3.9990091651326829E-5, -4.0090852176581095E-5, -4.0154101038240283E-5, -4.0181466434390562E-5, -4.017453316660271E-5, -4.013484327935801E-5, -4.0063896706025282E-5, -3.9963151920563813E-5, -3.9834026594159355E-5, -3.9677898256031791E-5, -3.9496104957683613E-5, -3.9289945939888413E-5, -3.9060682301747689E-5, -3.8809537671172525E-5, -3.8537698876174604E-5, -3.8246316616377579E-5, -3.793650613418646E-5, -3.7609347885077623E-5, -3.7265888206497395E-5, -3.6907139984880808E-5, -3.6534083320325723E-5, -3.6147666188480321E-5, -3.5748805099224027E-5, -3.5338385751743129E-5, -3.4917263685623729E-5, -3.44862649276042E-5, -3.40461866336495E-5, -3.3597797726028135E-5, -3.3141839525091535E-5, -3.2679026375472935E-5, -3.221004626644033E-5, -3.1735561446154833E-5, -3.12562090296018E-5, -3.0772601599977736E-5, -3.0285327803331116E-5, -2.9794952936269942E-5, -2.9302019526562752E-5, -2.8807047906473585E-5, -2.8310536778684464E-5, -2.7812963774671571E-5, -2.7314786005413577E-5, -2.6816440604322343E-5, -2.6318345262297408E-5, -2.5820898754816765E-5, -2.5324481460986734E-5, -2.4829455874483883E-5, -2.4336167106331684E-5, -2.3844943379463754E-5, -2.3356096515034559E-5, -2.2869922410446928E-5, -2.2386701509073987E-5, -2.190669926166088E-5, -2.1430166579399207E-5, -2.0957340278674263E-5, -2.0488443517492027E-5, -2.0023686223599328E-5, -1.9563265514316956E-5, -1.910736610811127E-5, -1.8656160727935741E-5, -1.8209810496378919E-5, -1.776846532266075E-5, -1.7332264281523728E-5, -1.6901335984070202E-5, -1.6475798940601218E-5, -1.6055761915516631E-5, -1.5641324274339943E-5, -1.5232576322934952E-5, -1.4829599638984815E-5, -1.4432467395807249E-5, -1.4041244678582621E-5, -1.3655988793074526E-5, -1.3276749566924981E-5, -1.29035696436089E-5, -1.2536484769134677E-5, -1.217552407157984E-5, -1.1820710333552607E-5, -1.1472060257671982E-5, -1.1129584725160594E-5, -1.0793289047645905E-5, -1.0463173212266783E-5, -1.0139232120183559E-5, -9.8214558185907186E-6, -9.5098297263323067E-6, -9.20433485322091E-6, -8.9049480131616991E-6, -8.6116420311836354E-6, -8.324385944480339E-6, -8.04314519756346E-6, -7.7678818316316609E-6, 0.0, 0.0, 0.0, 0.0, 0.0, 1.7756006070928429E-5, 1.955926027849794E-5, 2.1265642444599059E-5, 2.2878087249309936E-5, 2.4399475238503513E-5, 2.5832632877734329E-5, 2.7180332648224444E-5, 2.8445293182983732E-5, 2.9630179441154765E-5, 3.0737602918726609E-5, 3.1770121893815045E-5, 3.2730241704758869E-5, 3.3620415059333691E-5, 3.4443042373434618E-5, 3.5200472137629193E-5, 3.5895001310030509E-5, 3.652887573398812E-5, 3.7104290579141277E-5, 3.7623390804425058E-5, 3.808827164166491E-5, 3.8500979098439383E-5, 3.886351047893401E-5, 3.9177814921551905E-5, 3.9445793952087749E-5, 3.966930205131298E-5, 3.98501472358593E-5, 3.9990091651326829E-5, 4.0090852176581095E-5, 4.0154101038240283E-5, 4.0181466434390562E-5, 4.017453316660271E-5, 4.013484327935801E-5, 4.0063896706025282E-5, 3.9963151920563813E-5, 3.9834026594159355E-5, 3.9677898256031791E-5, 3.9496104957683613E-5, 3.9289945939888413E-5, 3.9060682301747689E-5, 3.8809537671172525E-5, 3.8537698876174604E-5, 3.8246316616377579E-5, 3.793650613418646E-5, 3.7609347885077623E-5, 3.7265888206497395E-5, 3.6907139984880808E-5, 3.6534083320325723E-5, 3.6147666188480321E-5, 3.5748805099224027E-5, 3.5338385751743129E-5, 3.4917263685623729E-5, 3.44862649276042E-5, 3.40461866336495E-5, 3.3597797726028135E-5, 3.3141839525091535E-5, 3.2679026375472935E-5, 3.221004626644033E-5, 3.1735561446154833E-5, 3.12562090296018E-5, 3.0772601599977736E-5, 3.0285327803331116E-5, 2.9794952936269942E-5, 2.9302019526562752E-5, 2.8807047906473585E-5, 2.8310536778684464E-5, 2.7812963774671571E-5, 2.7314786005413577E-5, 2.6816440604322343E-5, 2.6318345262297408E-5, 2.5820898754816765E-5, 2.5324481460986734E-5, 2.4829455874483883E-5, 2.4336167106331684E-5, 2.3844943379463754E-5, 2.3356096515034559E-5, 2.2869922410446928E-5, 2.2386701509073987E-5, 2.190669926166088E-5, 2.1430166579399207E-5, 2.0957340278674263E-5, 2.0488443517492027E-5, 2.0023686223599328E-5, 1.9563265514316956E-5, 1.910736610811127E-5, 1.8656160727935741E-5, 1.8209810496378919E-5, 1.776846532266075E-5, 1.7332264281523728E-5, 1.6901335984070202E-5, 1.6475798940601218E-5, 1.6055761915516631E-5, 1.5641324274339943E-5, 1.5232576322934952E-5, 1.4829599638984815E-5, 1.4432467395807249E-5, 1.4041244678582621E-5, 1.3655988793074526E-5, 1.3276749566924981E-5, 1.29035696436089E-5, 1.2536484769134677E-5, 1.217552407157984E-5, 1.1820710333552607E-5, 1.1472060257671982E-5, 1.1129584725160594E-5, 1.0793289047645905E-5, 1.0463173212266783E-5, 1.0139232120183559E-5, 9.8214558185907186E-6, 9.5098297263323067E-6, 9.20433485322091E-6, 8.9049480131616991E-6, 8.6116420311836354E-6, 8.324385944480339E-6, 8.04314519756346E-6, 7.7678818316316609E-6, 0.0, 0.0, 0.0, 0.0, -0.0, -0.0, -0.0, -0.0, -0.0, -0.0, -0.0, -0.0, -0.0, -0.0, -0.0, -0.0, -0.0, -0.0, -0.0, -0.0, -0.0, -0.0, -0.0, -0.0, -0.0, -0.0, -0.0, -0.0, -0.0, -0.0, -0.0, -0.0, -0.0, -0.0, -0.0, -0.0, -0.0, -0.0, -0.0, -0.0, -0.0, -0.0, -0.0, -0.0, -0.0, -0.0, -0.0, -0.0, -0.0, -0.0, -0.0, -0.0, -0.0, -0.0, -0.0, -0.0, -0.0, -0.0, -0.0, -0.0, -0.0, -0.0, -0.0, -0.0, -0.0, -0.0, -0.0, -0.0, -0.0, -0.0, -0.0, -0.0, -0.0, -0.0, -0.0, -0.0, -0.0, -0.0, -0.0, -0.0, -0.0, -0.0, -0.0, -0.0, -0.0, -0.0, -0.0, -0.0, -0.0, -0.0, -0.0, -0.0, -0.0, -0.0, -0.0, -0.0, -0.0, -0.0, -0.0, -0.0, -0.0, -0.0, -0.0, -0.0, -0.0, -0.0, -0.0, -0.0, -0.0, -0.0, -0.0, -0.0, -0.0, -0.0, -0.0, -0.0, -0.0, -0.0, -0.0, -0.0, -0.0, -0.0, -0.0, -0.0, 0.0, 0.0, 0.0, 0.0, 0.0, 0.0, 0.0, 0.0, 0.0, 0.0, 0.0, 0.0, 0.0, 0.0, 0.0, 0.0, 0.0, 0.0, 0.0, 0.0, 0.0, 0.0, 0.0, 0.0, 0.0, 0.0, 0.0, 0.0, 0.0, 0.0, 0.0, 0.0, 0.0, 0.0, 0.0, 0.0, 0.0, 0.0, 0.0, 0.0, 0.0, 0.0, 0.0, 0.0, 0.0, 0.0, 0.0, 0.0, 0.0, 0.0, 0.0, 0.0, 0.0, 0.0, 0.0, 0.0, 0.0, 0.0, 0.0, 0.0, 0.0, 0.0, 0.0, 0.0, 0.0, 0.0, 0.0, 0.0, 0.0, 0.0, 0.0, 0.0, 0.0, 0.0, 0.0, 0.0, 0.0, 0.0, 0.0, 0.0, 0.0, 0.0, 0.0, 0.0, 0.0, 0.0, 0.0, 0.0, 0.0, 0.0, 0.0, 0.0, 0.0, 0.0, 0.0, 0.0, 0.0, 0.0, 0.0, 0.0, 0.0, 0.0, 0.0, 0.0, 0.0, 0.0, 0.0, 0.0, 0.0, 0.0, 0.0, 0.0, 0.0, 0.0, 0.0, 0.0, 0.0, 0.0, 0.0, 0.0, 0.0, 0.0, 0.0, 0.0, -0.0, -0.0, -0.0, -0.0, -0.0, -0.0, -1.7756006070928429E-5, -1.955926027849794E-5, -2.1265642444599059E-5, -2.2878087249309936E-5, -2.4399475238503513E-5, -2.5832632877734329E-5, -2.7180332648224444E-5, -2.8445293182983732E-5, -2.9630179441154765E-5, -3.0737602918726609E-5, -3.1770121893815045E-5, -3.2730241704758869E-5, -3.3620415059333691E-5, -3.4443042373434618E-5, -3.5200472137629193E-5, -3.5895001310030509E-5, -3.652887573398812E-5, -3.7104290579141277E-5, -3.7623390804425058E-5, -3.808827164166491E-5, -3.8500979098439383E-5, -3.886351047893401E-5, -3.9177814921551905E-5, -3.9445793952087749E-5, -3.966930205131298E-5, -3.98501472358593E-5, -3.9990091651326829E-5, -4.0090852176581095E-5, -4.0154101038240283E-5, -4.0181466434390562E-5, -4.017453316660271E-5, -4.013484327935801E-5, -4.0063896706025282E-5, -3.9963151920563813E-5, -3.9834026594159355E-5, -3.9677898256031791E-5, -3.9496104957683613E-5, -3.9289945939888413E-5, -3.9060682301747689E-5, -3.8809537671172525E-5, -3.8537698876174604E-5, -3.8246316616377579E-5, -3.793650613418646E-5, -3.7609347885077623E-5, -3.7265888206497395E-5, -3.6907139984880808E-5, -3.6534083320325723E-5, -3.6147666188480321E-5, -3.5748805099224027E-5, -3.5338385751743129E-5, -3.4917263685623729E-5, -3.44862649276042E-5, -3.40461866336495E-5, -3.3597797726028135E-5, -3.3141839525091535E-5, -3.2679026375472935E-5, -3.221004626644033E-5, -3.1735561446154833E-5, -3.12562090296018E-5, -3.0772601599977736E-5, -3.0285327803331116E-5, -2.9794952936269942E-5, -2.9302019526562752E-5, -2.8807047906473585E-5, -2.8310536778684464E-5, -2.7812963774671571E-5, -2.7314786005413577E-5, -2.6816440604322343E-5, -2.6318345262297408E-5, -2.5820898754816765E-5, -2.5324481460986734E-5, -2.4829455874483883E-5, -2.4336167106331684E-5, -2.3844943379463754E-5, -2.3356096515034559E-5, -2.2869922410446928E-5, -2.2386701509073987E-5, -2.190669926166088E-5, -2.1430166579399207E-5, -2.0957340278674263E-5, -2.0488443517492027E-5, -2.0023686223599328E-5, -1.9563265514316956E-5, -1.910736610811127E-5, -1.8656160727935741E-5, -1.8209810496378919E-5, -1.776846532266075E-5, -1.7332264281523728E-5, -1.6901335984070202E-5, -1.6475798940601218E-5, -1.6055761915516631E-5, -1.5641324274339943E-5, -1.5232576322934952E-5, -1.4829599638984815E-5, -1.4432467395807249E-5, -1.4041244678582621E-5, -1.3655988793074526E-5, -1.3276749566924981E-5, -1.29035696436089E-5, -1.2536484769134677E-5, -1.217552407157984E-5, -1.1820710333552607E-5, -1.1472060257671982E-5, -1.1129584725160594E-5, -1.0793289047645905E-5, -1.0463173212266783E-5, -1.0139232120183559E-5, -9.8214558185907186E-6, -9.5098297263323067E-6, -9.20433485322091E-6, -8.9049480131616991E-6, -8.6116420311836354E-6, -8.324385944480339E-6, -8.04314519756346E-6, 0.0, 0.0, 0.0, 0.0, 0.0, 0.0, 1.7756006070928429E-5, 1.955926027849794E-5, 2.1265642444599059E-5, 2.2878087249309936E-5, 2.4399475238503513E-5, 2.5832632877734329E-5, 2.7180332648224444E-5, 2.8445293182983732E-5, 2.9630179441154765E-5, 3.0737602918726609E-5, 3.1770121893815045E-5, 3.2730241704758869E-5, 3.3620415059333691E-5, 3.4443042373434618E-5, 3.5200472137629193E-5, 3.5895001310030509E-5, 3.652887573398812E-5, 3.7104290579141277E-5, 3.7623390804425058E-5, 3.808827164166491E-5, 3.8500979098439383E-5, 3.886351047893401E-5, 3.9177814921551905E-5, 3.9445793952087749E-5, 3.966930205131298E-5, 3.98501472358593E-5, 3.9990091651326829E-5, 4.0090852176581095E-5, 4.0154101038240283E-5, 4.0181466434390562E-5, 4.017453316660271E-5, 4.013484327935801E-5, 4.0063896706025282E-5, 3.9963151920563813E-5, 3.9834026594159355E-5, 3.9677898256031791E-5, 3.9496104957683613E-5, 3.9289945939888413E-5, 3.9060682301747689E-5, 3.8809537671172525E-5, 3.8537698876174604E-5, 3.8246316616377579E-5, 3.793650613418646E-5, 3.7609347885077623E-5, 3.7265888206497395E-5, 3.6907139984880808E-5, 3.6534083320325723E-5, 3.6147666188480321E-5, 3.5748805099224027E-5, 3.5338385751743129E-5, 3.4917263685623729E-5, 3.44862649276042E-5, 3.40461866336495E-5, 3.3597797726028135E-5, 3.3141839525091535E-5, 3.2679026375472935E-5, 3.221004626644033E-5, 3.1735561446154833E-5, 3.12562090296018E-5, 3.0772601599977736E-5, 3.0285327803331116E-5, 2.9794952936269942E-5, 2.9302019526562752E-5, 2.8807047906473585E-5, 2.8310536778684464E-5, 2.7812963774671571E-5, 2.7314786005413577E-5, 2.6816440604322343E-5, 2.6318345262297408E-5, 2.5820898754816765E-5, 2.5324481460986734E-5, 2.4829455874483883E-5, 2.4336167106331684E-5, 2.3844943379463754E-5, 2.3356096515034559E-5, 2.2869922410446928E-5, 2.2386701509073987E-5, 2.190669926166088E-5, 2.1430166579399207E-5, 2.0957340278674263E-5, 2.0488443517492027E-5, 2.0023686223599328E-5, 1.9563265514316956E-5, 1.910736610811127E-5, 1.8656160727935741E-5, 1.8209810496378919E-5, 1.776846532266075E-5, 1.7332264281523728E-5, 1.6901335984070202E-5, 1.6475798940601218E-5, 1.6055761915516631E-5, 1.5641324274339943E-5, 1.5232576322934952E-5, 1.4829599638984815E-5, 1.4432467395807249E-5, 1.4041244678582621E-5, 1.3655988793074526E-5, 1.3276749566924981E-5, 1.29035696436089E-5, 1.2536484769134677E-5, 1.217552407157984E-5, 1.1820710333552607E-5, 1.1472060257671982E-5, 1.1129584725160594E-5, 1.0793289047645905E-5, 1.0463173212266783E-5, 1.0139232120183559E-5, 9.8214558185907186E-6, 9.5098297263323067E-6, 9.20433485322091E-6, 8.9049480131616991E-6, 8.6116420311836354E-6, 8.324385944480339E-6, 8.04314519756346E-6, 0.0, 0.0, 0.0, 0.0, -0.0, -0.0, -0.0, -0.0, -0.0, -0.0, -0.0, -0.0, -0.0, -0.0, -0.0, -0.0, -0.0, -0.0, -0.0, -0.0, -0.0, -0.0, -0.0, -0.0, -0.0, -0.0, -0.0, -0.0, -0.0, -0.0, -0.0, -0.0, -0.0, -0.0, -0.0, -0.0, -0.0, -0.0, -0.0, -0.0, -0.0, -0.0, -0.0, -0.0, -0.0, -0.0, -0.0, -0.0, -0.0, -0.0, -0.0, -0.0, -0.0, -0.0, -0.0, -0.0, -0.0, -0.0, -0.0, -0.0, -0.0, -0.0, -0.0, -0.0, -0.0, -0.0, -0.0, -0.0, -0.0, -0.0, -0.0, -0.0, -0.0, -0.0, -0.0, -0.0, -0.0, -0.0, -0.0, -0.0, -0.0, -0.0, -0.0, -0.0, -0.0, -0.0, -0.0, -0.0, -0.0, -0.0, -0.0, -0.0, -0.0, -0.0, -0.0, -0.0, -0.0, -0.0, -0.0, -0.0, -0.0, -0.0, -0.0, -0.0, -0.0, -0.0, -0.0, -0.0, -0.0, -0.0, -0.0, -0.0, -0.0, -0.0, -0.0, -0.0, -0.0, -0.0, -0.0, -0.0, -0.0, -0.0, -0.0, -0.0, 0.0, 0.0, 0.0, 0.0, 0.0, 0.0, 0.0, 0.0, 0.0, 0.0, 0.0, 0.0, 0.0, 0.0, 0.0, 0.0, 0.0, 0.0, 0.0, 0.0, 0.0, 0.0, 0.0, 0.0, 0.0, 0.0, 0.0, 0.0, 0.0, 0.0, 0.0, 0.0, 0.0, 0.0, 0.0, 0.0, 0.0, 0.0, 0.0, 0.0, 0.0, 0.0, 0.0, 0.0, 0.0, 0.0, 0.0, 0.0, 0.0, 0.0, 0.0, 0.0, 0.0, 0.0, 0.0, 0.0, 0.0, 0.0, 0.0, 0.0, 0.0, 0.0, 0.0, 0.0, 0.0, 0.0, 0.0, 0.0, 0.0, 0.0, 0.0, 0.0, 0.0, 0.0, 0.0, 0.0, 0.0, 0.0, 0.0, 0.0, 0.0, 0.0, 0.0, 0.0, 0.0, 0.0, 0.0, 0.0, 0.0, 0.0, 0.0, 0.0, 0.0, 0.0, 0.0, 0.0, 0.0, 0.0, 0.0, 0.0, 0.0, 0.0, 0.0, 0.0, 0.0, 0.0, 0.0, 0.0, 0.0, 0.0, 0.0, 0.0, 0.0, 0.0, 0.0, 0.0, 0.0, 0.0, 0.0, 0.0, 0.0, 0.0, 0.0, 0.0, -0.0, -0.0, -0.0, -0.0, -0.0, -0.0, -0.0, -1.7756006070928429E-5, -1.955926027849794E-5, -2.1265642444599059E-5, -2.2878087249309936E-5, -2.4399475238503513E-5, -2.5832632877734329E-5, -2.7180332648224444E-5, -2.8445293182983732E-5, -2.9630179441154765E-5, -3.0737602918726609E-5, -3.1770121893815045E-5, -3.2730241704758869E-5, -3.3620415059333691E-5, -3.4443042373434618E-5, -3.5200472137629193E-5, -3.5895001310030509E-5, -3.652887573398812E-5, -3.7104290579141277E-5, -3.7623390804425058E-5, -3.808827164166491E-5, -3.8500979098439383E-5, -3.886351047893401E-5, -3.9177814921551905E-5, -3.9445793952087749E-5, -3.966930205131298E-5, -3.98501472358593E-5, -3.9990091651326829E-5, -4.0090852176581095E-5, -4.0154101038240283E-5, -4.0181466434390562E-5, -4.017453316660271E-5, -4.013484327935801E-5, -4.0063896706025282E-5, -3.9963151920563813E-5, -3.9834026594159355E-5, -3.9677898256031791E-5, -3.9496104957683613E-5, -3.9289945939888413E-5, -3.9060682301747689E-5, -3.8809537671172525E-5, -3.8537698876174604E-5, -3.8246316616377579E-5, -3.793650613418646E-5, -3.7609347885077623E-5, -3.7265888206497395E-5, -3.6907139984880808E-5, -3.6534083320325723E-5, -3.6147666188480321E-5, -3.5748805099224027E-5, -3.5338385751743129E-5, -3.4917263685623729E-5, -3.44862649276042E-5, -3.40461866336495E-5, -3.3597797726028135E-5, -3.3141839525091535E-5, -3.2679026375472935E-5, -3.221004626644033E-5, -3.1735561446154833E-5, -3.12562090296018E-5, -3.0772601599977736E-5, -3.0285327803331116E-5, -2.9794952936269942E-5, -2.9302019526562752E-5, -2.8807047906473585E-5, -2.8310536778684464E-5, -2.7812963774671571E-5, -2.7314786005413577E-5, -2.6816440604322343E-5, -2.6318345262297408E-5, -2.5820898754816765E-5, -2.5324481460986734E-5, -2.4829455874483883E-5, -2.4336167106331684E-5, -2.3844943379463754E-5, -2.3356096515034559E-5, -2.2869922410446928E-5, -2.2386701509073987E-5, -2.190669926166088E-5, -2.1430166579399207E-5, -2.0957340278674263E-5, -2.0488443517492027E-5, -2.0023686223599328E-5, -1.9563265514316956E-5, -1.910736610811127E-5, -1.8656160727935741E-5, -1.8209810496378919E-5, -1.776846532266075E-5, -1.7332264281523728E-5, -1.6901335984070202E-5, -1.6475798940601218E-5, -1.6055761915516631E-5, -1.5641324274339943E-5, -1.5232576322934952E-5, -1.4829599638984815E-5, -1.4432467395807249E-5, -1.4041244678582621E-5, -1.3655988793074526E-5, -1.3276749566924981E-5, -1.29035696436089E-5, -1.2536484769134677E-5, -1.217552407157984E-5, -1.1820710333552607E-5, -1.1472060257671982E-5, -1.1129584725160594E-5, -1.0793289047645905E-5, -1.0463173212266783E-5, -1.0139232120183559E-5, -9.8214558185907186E-6, -9.5098297263323067E-6, -9.20433485322091E-6, -8.9049480131616991E-6, -8.6116420311836354E-6, -8.324385944480339E-6, 0.0, 0.0, 0.0, 0.0, 0.0, 0.0, 0.0, 1.7756006070928429E-5, 1.955926027849794E-5, 2.1265642444599059E-5, 2.2878087249309936E-5, 2.4399475238503513E-5, 2.5832632877734329E-5, 2.7180332648224444E-5, 2.8445293182983732E-5, 2.9630179441154765E-5, 3.0737602918726609E-5, 3.1770121893815045E-5, 3.2730241704758869E-5, 3.3620415059333691E-5, 3.4443042373434618E-5, 3.5200472137629193E-5, 3.5895001310030509E-5, 3.652887573398812E-5, 3.7104290579141277E-5, 3.7623390804425058E-5, 3.808827164166491E-5, 3.8500979098439383E-5, 3.886351047893401E-5, 3.9177814921551905E-5, 3.9445793952087749E-5, 3.966930205131298E-5, 3.98501472358593E-5, 3.9990091651326829E-5, 4.0090852176581095E-5, 4.0154101038240283E-5, 4.0181466434390562E-5, 4.017453316660271E-5, 4.013484327935801E-5, 4.0063896706025282E-5, 3.9963151920563813E-5, 3.9834026594159355E-5, 3.9677898256031791E-5, 3.9496104957683613E-5, 3.9289945939888413E-5, 3.9060682301747689E-5, 3.8809537671172525E-5, 3.8537698876174604E-5, 3.8246316616377579E-5, 3.793650613418646E-5, 3.7609347885077623E-5, 3.7265888206497395E-5, 3.6907139984880808E-5, 3.6534083320325723E-5, 3.6147666188480321E-5, 3.5748805099224027E-5, 3.5338385751743129E-5, 3.4917263685623729E-5, 3.44862649276042E-5, 3.40461866336495E-5, 3.3597797726028135E-5, 3.3141839525091535E-5, 3.2679026375472935E-5, 3.221004626644033E-5, 3.1735561446154833E-5, 3.12562090296018E-5, 3.0772601599977736E-5, 3.0285327803331116E-5, 2.9794952936269942E-5, 2.9302019526562752E-5, 2.8807047906473585E-5, 2.8310536778684464E-5, 2.7812963774671571E-5, 2.7314786005413577E-5, 2.6816440604322343E-5, 2.6318345262297408E-5, 2.5820898754816765E-5, 2.5324481460986734E-5, 2.4829455874483883E-5, 2.4336167106331684E-5, 2.3844943379463754E-5, 2.3356096515034559E-5, 2.2869922410446928E-5, 2.2386701509073987E-5, 2.190669926166088E-5, 2.1430166579399207E-5, 2.0957340278674263E-5, 2.0488443517492027E-5, 2.0023686223599328E-5, 1.9563265514316956E-5, 1.910736610811127E-5, 1.8656160727935741E-5, 1.8209810496378919E-5, 1.776846532266075E-5, 1.7332264281523728E-5, 1.6901335984070202E-5, 1.6475798940601218E-5, 1.6055761915516631E-5, 1.5641324274339943E-5, 1.5232576322934952E-5, 1.4829599638984815E-5, 1.4432467395807249E-5, 1.4041244678582621E-5, 1.3655988793074526E-5, 1.3276749566924981E-5, 1.29035696436089E-5, 1.2536484769134677E-5, 1.217552407157984E-5, 1.1820710333552607E-5, 1.1472060257671982E-5, 1.1129584725160594E-5, 1.0793289047645905E-5, 1.0463173212266783E-5, 1.0139232120183559E-5, 9.8214558185907186E-6, 9.5098297263323067E-6, 9.20433485322091E-6, 8.9049480131616991E-6, 8.6116420311836354E-6, 8.324385944480339E-6, 0.0, 0.0, 0.0, 0.0, -0.0, -0.0, -0.0, -0.0, -0.0, -0.0, -0.0, -0.0, -0.0, -0.0, -0.0, -0.0, -0.0, -0.0, -0.0, -0.0, -0.0, -0.0, -0.0, -0.0, -0.0, -0.0, -0.0, -0.0, -0.0, -0.0, -0.0, -0.0, -0.0, -0.0, -0.0, -0.0, -0.0, -0.0, -0.0, -0.0, -0.0, -0.0, -0.0, -0.0, -0.0, -0.0, -0.0, -0.0, -0.0, -0.0, -0.0, -0.0, -0.0, -0.0, -0.0, -0.0, -0.0, -0.0, -0.0, -0.0, -0.0, -0.0, -0.0, -0.0, -0.0, -0.0, -0.0, -0.0, -0.0, -0.0, -0.0, -0.0, -0.0, -0.0, -0.0, -0.0, -0.0, -0.0, -0.0, -0.0, -0.0, -0.0, -0.0, -0.0, -0.0, -0.0, -0.0, -0.0, -0.0, -0.0, -0.0, -0.0, -0.0, -0.0, -0.0, -0.0, -0.0, -0.0, -0.0, -0.0, -0.0, -0.0, -0.0, -0.0, -0.0, -0.0, -0.0, -0.0, -0.0, -0.0, -0.0, -0.0, -0.0, -0.0, -0.0, -0.0, -0.0, -0.0, -0.0, -0.0, -0.0, -0.0, -0.0, -0.0, 0.0, 0.0, 0.0, 0.0, 0.0, 0.0, 0.0, 0.0, 0.0, 0.0, 0.0, 0.0, 0.0, 0.0, 0.0, 0.0, 0.0, 0.0, 0.0, 0.0, 0.0, 0.0, 0.0, 0.0, 0.0, 0.0, 0.0, 0.0, 0.0, 0.0, 0.0, 0.0, 0.0, 0.0, 0.0, 0.0, 0.0, 0.0, 0.0, 0.0, 0.0, 0.0, 0.0, 0.0, 0.0, 0.0, 0.0, 0.0, 0.0, 0.0, 0.0, 0.0, 0.0, 0.0, 0.0, 0.0, 0.0, 0.0, 0.0, 0.0, 0.0, 0.0, 0.0, 0.0, 0.0, 0.0, 0.0, 0.0, 0.0, 0.0, 0.0, 0.0, 0.0, 0.0, 0.0, 0.0, 0.0, 0.0, 0.0, 0.0, 0.0, 0.0, 0.0, 0.0, 0.0, 0.0, 0.0, 0.0, 0.0, 0.0, 0.0, 0.0, 0.0, 0.0, 0.0, 0.0, 0.0, 0.0, 0.0, 0.0, 0.0, 0.0, 0.0, 0.0, 0.0, 0.0, 0.0, 0.0, 0.0, 0.0, 0.0, 0.0, 0.0, 0.0, 0.0, 0.0, 0.0, 0.0, 0.0, 0.0, 0.0, 0.0, 0.0, 0.0, -0.0, -0.0, -0.0, -0.0, -0.0, -0.0, -0.0, -0.0, -1.7756006070928429E-5, -1.955926027849794E-5, -2.1265642444599059E-5, -2.2878087249309936E-5, -2.4399475238503513E-5, -2.5832632877734329E-5, -2.7180332648224444E-5, -2.8445293182983732E-5, -2.9630179441154765E-5, -3.0737602918726609E-5, -3.1770121893815045E-5, -3.2730241704758869E-5, -3.3620415059333691E-5, -3.4443042373434618E-5, -3.5200472137629193E-5, -3.5895001310030509E-5, -3.652887573398812E-5, -3.7104290579141277E-5, -3.7623390804425058E-5, -3.808827164166491E-5, -3.8500979098439383E-5, -3.886351047893401E-5, -3.9177814921551905E-5, -3.9445793952087749E-5, -3.966930205131298E-5, -3.98501472358593E-5, -3.9990091651326829E-5, -4.0090852176581095E-5, -4.0154101038240283E-5, -4.0181466434390562E-5, -4.017453316660271E-5, -4.013484327935801E-5, -4.0063896706025282E-5, -3.9963151920563813E-5, -3.9834026594159355E-5, -3.9677898256031791E-5, -3.9496104957683613E-5, -3.9289945939888413E-5, -3.9060682301747689E-5, -3.8809537671172525E-5, -3.8537698876174604E-5, -3.8246316616377579E-5, -3.793650613418646E-5, -3.7609347885077623E-5, -3.7265888206497395E-5, -3.6907139984880808E-5, -3.6534083320325723E-5, -3.6147666188480321E-5, -3.5748805099224027E-5, -3.5338385751743129E-5, -3.4917263685623729E-5, -3.44862649276042E-5, -3.40461866336495E-5, -3.3597797726028135E-5, -3.3141839525091535E-5, -3.2679026375472935E-5, -3.221004626644033E-5, -3.1735561446154833E-5, -3.12562090296018E-5, -3.0772601599977736E-5, -3.0285327803331116E-5, -2.9794952936269942E-5, -2.9302019526562752E-5, -2.8807047906473585E-5, -2.8310536778684464E-5, -2.7812963774671571E-5, -2.7314786005413577E-5, -2.6816440604322343E-5, -2.6318345262297408E-5, -2.5820898754816765E-5, -2.5324481460986734E-5, -2.4829455874483883E-5, -2.4336167106331684E-5, -2.3844943379463754E-5, -2.3356096515034559E-5, -2.2869922410446928E-5, -2.2386701509073987E-5, -2.190669926166088E-5, -2.1430166579399207E-5, -2.0957340278674263E-5, -2.0488443517492027E-5, -2.0023686223599328E-5, -1.9563265514316956E-5, -1.910736610811127E-5, -1.8656160727935741E-5, -1.8209810496378919E-5, -1.776846532266075E-5, -1.7332264281523728E-5, -1.6901335984070202E-5, -1.6475798940601218E-5, -1.6055761915516631E-5, -1.5641324274339943E-5, -1.5232576322934952E-5, -1.4829599638984815E-5, -1.4432467395807249E-5, -1.4041244678582621E-5, -1.3655988793074526E-5, -1.3276749566924981E-5, -1.29035696436089E-5, -1.2536484769134677E-5, -1.217552407157984E-5, -1.1820710333552607E-5, -1.1472060257671982E-5, -1.1129584725160594E-5, -1.0793289047645905E-5, -1.0463173212266783E-5, -1.0139232120183559E-5, -9.8214558185907186E-6, -9.5098297263323067E-6, -9.20433485322091E-6, -8.9049480131616991E-6, -8.6116420311836354E-6, 0.0, 0.0, 0.0, 0.0, 0.0, 0.0, 0.0, 0.0, 1.7756006070928429E-5, 1.955926027849794E-5, 2.1265642444599059E-5, 2.2878087249309936E-5, 2.4399475238503513E-5, 2.5832632877734329E-5, 2.7180332648224444E-5, 2.8445293182983732E-5, 2.9630179441154765E-5, 3.0737602918726609E-5, 3.1770121893815045E-5, 3.2730241704758869E-5, 3.3620415059333691E-5, 3.4443042373434618E-5, 3.5200472137629193E-5, 3.5895001310030509E-5, 3.652887573398812E-5, 3.7104290579141277E-5, 3.7623390804425058E-5, 3.808827164166491E-5, 3.8500979098439383E-5, 3.886351047893401E-5, 3.9177814921551905E-5, 3.9445793952087749E-5, 3.966930205131298E-5, 3.98501472358593E-5, 3.9990091651326829E-5, 4.0090852176581095E-5, 4.0154101038240283E-5, 4.0181466434390562E-5, 4.017453316660271E-5, 4.013484327935801E-5, 4.0063896706025282E-5, 3.9963151920563813E-5, 3.9834026594159355E-5, 3.9677898256031791E-5, 3.9496104957683613E-5, 3.9289945939888413E-5, 3.9060682301747689E-5, 3.8809537671172525E-5, 3.8537698876174604E-5, 3.8246316616377579E-5, 3.793650613418646E-5, 3.7609347885077623E-5, 3.7265888206497395E-5, 3.6907139984880808E-5, 3.6534083320325723E-5, 3.6147666188480321E-5, 3.5748805099224027E-5, 3.5338385751743129E-5, 3.4917263685623729E-5, 3.44862649276042E-5, 3.40461866336495E-5, 3.3597797726028135E-5, 3.3141839525091535E-5, 3.2679026375472935E-5, 3.221004626644033E-5, 3.1735561446154833E-5, 3.12562090296018E-5, 3.0772601599977736E-5, 3.0285327803331116E-5, 2.9794952936269942E-5, 2.9302019526562752E-5, 2.8807047906473585E-5, 2.8310536778684464E-5, 2.7812963774671571E-5, 2.7314786005413577E-5, 2.6816440604322343E-5, 2.6318345262297408E-5, 2.5820898754816765E-5, 2.5324481460986734E-5, 2.4829455874483883E-5, 2.4336167106331684E-5, 2.3844943379463754E-5, 2.3356096515034559E-5, 2.2869922410446928E-5, 2.2386701509073987E-5, 2.190669926166088E-5, 2.1430166579399207E-5, 2.0957340278674263E-5, 2.0488443517492027E-5, 2.0023686223599328E-5, 1.9563265514316956E-5, 1.910736610811127E-5, 1.8656160727935741E-5, 1.8209810496378919E-5, 1.776846532266075E-5, 1.7332264281523728E-5, 1.6901335984070202E-5, 1.6475798940601218E-5, 1.6055761915516631E-5, 1.5641324274339943E-5, 1.5232576322934952E-5, 1.4829599638984815E-5, 1.4432467395807249E-5, 1.4041244678582621E-5, 1.3655988793074526E-5, 1.3276749566924981E-5, 1.29035696436089E-5, 1.2536484769134677E-5, 1.217552407157984E-5, 1.1820710333552607E-5, 1.1472060257671982E-5, 1.1129584725160594E-5, 1.0793289047645905E-5, 1.0463173212266783E-5, 1.0139232120183559E-5, 9.8214558185907186E-6, 9.5098297263323067E-6, 9.20433485322091E-6, 8.9049480131616991E-6, 8.6116420311836354E-6, 0.0, 0.0, 0.0, 0.0, -0.0, -0.0, -0.0, -0.0, -0.0, -0.0, -0.0, -0.0, -0.0, -0.0, -0.0, -0.0, -0.0, -0.0, -0.0, -0.0, -0.0, -0.0, -0.0, -0.0, -0.0, -0.0, -0.0, -0.0, -0.0, -0.0, -0.0, -0.0, -0.0, -0.0, -0.0, -0.0, -0.0, -0.0, -0.0, -0.0, -0.0, -0.0, -0.0, -0.0, -0.0, -0.0, -0.0, -0.0, -0.0, -0.0, -0.0, -0.0, -0.0, -0.0, -0.0, -0.0, -0.0, -0.0, -0.0, -0.0, -0.0, -0.0, -0.0, -0.0, -0.0, -0.0, -0.0, -0.0, -0.0, -0.0, -0.0, -0.0, -0.0, -0.0, -0.0, -0.0, -0.0, -0.0, -0.0, -0.0, -0.0, -0.0, -0.0, -0.0, -0.0, -0.0, -0.0, -0.0, -0.0, -0.0, -0.0, -0.0, -0.0, -0.0, -0.0, -0.0, -0.0, -0.0, -0.0, -0.0, -0.0, -0.0, -0.0, -0.0, -0.0, -0.0, -0.0, -0.0, -0.0, -0.0, -0.0, -0.0, -0.0, -0.0, -0.0, -0.0, -0.0, -0.0, -0.0, -0.0, -0.0, -0.0, -0.0, -0.0, 0.0, 0.0, 0.0, 0.0, 0.0, 0.0, 0.0, 0.0, 0.0, 0.0, 0.0, 0.0, 0.0, 0.0, 0.0, 0.0, 0.0, 0.0, 0.0, 0.0, 0.0, 0.0, 0.0, 0.0, 0.0, 0.0, 0.0, 0.0, 0.0, 0.0, 0.0, 0.0, 0.0, 0.0, 0.0, 0.0, 0.0, 0.0, 0.0, 0.0, 0.0, 0.0, 0.0, 0.0, 0.0, 0.0, 0.0, 0.0, 0.0, 0.0, 0.0, 0.0, 0.0, 0.0, 0.0, 0.0, 0.0, 0.0, 0.0, 0.0, 0.0, 0.0, 0.0, 0.0, 0.0, 0.0, 0.0, 0.0, 0.0, 0.0, 0.0, 0.0, 0.0, 0.0, 0.0, 0.0, 0.0, 0.0, 0.0, 0.0, 0.0, 0.0, 0.0, 0.0, 0.0, 0.0, 0.0, 0.0, 0.0, 0.0, 0.0, 0.0, 0.0, 0.0, 0.0, 0.0, 0.0, 0.0, 0.0, 0.0, 0.0, 0.0, 0.0, 0.0, 0.0, 0.0, 0.0, 0.0, 0.0, 0.0, 0.0, 0.0, 0.0, 0.0, 0.0, 0.0, 0.0, 0.0, 0.0, 0.0, 0.0, 0.0, 0.0, 0.0, -0.0, -0.0, -0.0, -0.0, -0.0, -0.0, -0.0, -0.0, -0.0, -1.7756006070928429E-5, -1.955926027849794E-5, -2.1265642444599059E-5, -2.2878087249309936E-5, -2.4399475238503513E-5, -2.5832632877734329E-5, -2.7180332648224444E-5, -2.8445293182983732E-5, -2.9630179441154765E-5, -3.0737602918726609E-5, -3.1770121893815045E-5, -3.2730241704758869E-5, -3.3620415059333691E-5, -3.4443042373434618E-5, -3.5200472137629193E-5, -3.5895001310030509E-5, -3.652887573398812E-5, -3.7104290579141277E-5, -3.7623390804425058E-5, -3.808827164166491E-5, -3.8500979098439383E-5, -3.886351047893401E-5, -3.9177814921551905E-5, -3.9445793952087749E-5, -3.966930205131298E-5, -3.98501472358593E-5, -3.9990091651326829E-5, -4.0090852176581095E-5, -4.0154101038240283E-5, -4.0181466434390562E-5, -4.017453316660271E-5, -4.013484327935801E-5, -4.0063896706025282E-5, -3.9963151920563813E-5, -3.9834026594159355E-5, -3.9677898256031791E-5, -3.9496104957683613E-5, -3.9289945939888413E-5, -3.9060682301747689E-5, -3.8809537671172525E-5, -3.8537698876174604E-5, -3.8246316616377579E-5, -3.793650613418646E-5, -3.7609347885077623E-5, -3.7265888206497395E-5, -3.6907139984880808E-5, -3.6534083320325723E-5, -3.6147666188480321E-5, -3.5748805099224027E-5, -3.5338385751743129E-5, -3.4917263685623729E-5, -3.44862649276042E-5, -3.40461866336495E-5, -3.3597797726028135E-5, -3.3141839525091535E-5, -3.2679026375472935E-5, -3.221004626644033E-5, -3.1735561446154833E-5, -3.12562090296018E-5, -3.0772601599977736E-5, -3.0285327803331116E-5, -2.9794952936269942E-5, -2.9302019526562752E-5, -2.8807047906473585E-5, -2.8310536778684464E-5, -2.7812963774671571E-5, -2.7314786005413577E-5, -2.6816440604322343E-5, -2.6318345262297408E-5, -2.5820898754816765E-5, -2.5324481460986734E-5, -2.4829455874483883E-5, -2.4336167106331684E-5, -2.3844943379463754E-5, -2.3356096515034559E-5, -2.2869922410446928E-5, -2.2386701509073987E-5, -2.190669926166088E-5, -2.1430166579399207E-5, -2.0957340278674263E-5, -2.0488443517492027E-5, -2.0023686223599328E-5, -1.9563265514316956E-5, -1.910736610811127E-5, -1.8656160727935741E-5, -1.8209810496378919E-5, -1.776846532266075E-5, -1.7332264281523728E-5, -1.6901335984070202E-5, -1.6475798940601218E-5, -1.6055761915516631E-5, -1.5641324274339943E-5, -1.5232576322934952E-5, -1.4829599638984815E-5, -1.4432467395807249E-5, -1.4041244678582621E-5, -1.3655988793074526E-5, -1.3276749566924981E-5, -1.29035696436089E-5, -1.2536484769134677E-5, -1.217552407157984E-5, -1.1820710333552607E-5, -1.1472060257671982E-5, -1.1129584725160594E-5, -1.0793289047645905E-5, -1.0463173212266783E-5, -1.0139232120183559E-5, -9.8214558185907186E-6, -9.5098297263323067E-6, -9.20433485322091E-6, -8.9049480131616991E-6, 0.0, 0.0, 0.0, 0.0, 0.0, 0.0, 0.0, 0.0, 0.0, 1.7756006070928429E-5, 1.955926027849794E-5, 2.1265642444599059E-5, 2.2878087249309936E-5, 2.4399475238503513E-5, 2.5832632877734329E-5, 2.7180332648224444E-5, 2.8445293182983732E-5, 2.9630179441154765E-5, 3.0737602918726609E-5, 3.1770121893815045E-5, 3.2730241704758869E-5, 3.3620415059333691E-5, 3.4443042373434618E-5, 3.5200472137629193E-5, 3.5895001310030509E-5, 3.652887573398812E-5, 3.7104290579141277E-5, 3.7623390804425058E-5, 3.808827164166491E-5, 3.8500979098439383E-5, 3.886351047893401E-5, 3.9177814921551905E-5, 3.9445793952087749E-5, 3.966930205131298E-5, 3.98501472358593E-5, 3.9990091651326829E-5, 4.0090852176581095E-5, 4.0154101038240283E-5, 4.0181466434390562E-5, 4.017453316660271E-5, 4.013484327935801E-5, 4.0063896706025282E-5, 3.9963151920563813E-5, 3.9834026594159355E-5, 3.9677898256031791E-5, 3.9496104957683613E-5, 3.9289945939888413E-5, 3.9060682301747689E-5, 3.8809537671172525E-5, 3.8537698876174604E-5, 3.8246316616377579E-5, 3.793650613418646E-5, 3.7609347885077623E-5, 3.7265888206497395E-5, 3.6907139984880808E-5, 3.6534083320325723E-5, 3.6147666188480321E-5, 3.5748805099224027E-5, 3.5338385751743129E-5, 3.4917263685623729E-5, 3.44862649276042E-5, 3.40461866336495E-5, 3.3597797726028135E-5, 3.3141839525091535E-5, 3.2679026375472935E-5, 3.221004626644033E-5, 3.1735561446154833E-5, 3.12562090296018E-5, 3.0772601599977736E-5, 3.0285327803331116E-5, 2.9794952936269942E-5, 2.9302019526562752E-5, 2.8807047906473585E-5, 2.8310536778684464E-5, 2.7812963774671571E-5, 2.7314786005413577E-5, 2.6816440604322343E-5, 2.6318345262297408E-5, 2.5820898754816765E-5, 2.5324481460986734E-5, 2.4829455874483883E-5, 2.4336167106331684E-5, 2.3844943379463754E-5, 2.3356096515034559E-5, 2.2869922410446928E-5, 2.2386701509073987E-5, 2.190669926166088E-5, 2.1430166579399207E-5, 2.0957340278674263E-5, 2.0488443517492027E-5, 2.0023686223599328E-5, 1.9563265514316956E-5, 1.910736610811127E-5, 1.8656160727935741E-5, 1.8209810496378919E-5, 1.776846532266075E-5, 1.7332264281523728E-5, 1.6901335984070202E-5, 1.6475798940601218E-5, 1.6055761915516631E-5, 1.5641324274339943E-5, 1.5232576322934952E-5, 1.4829599638984815E-5, 1.4432467395807249E-5, 1.4041244678582621E-5, 1.3655988793074526E-5, 1.3276749566924981E-5, 1.29035696436089E-5, 1.2536484769134677E-5, 1.217552407157984E-5, 1.1820710333552607E-5, 1.1472060257671982E-5, 1.1129584725160594E-5, 1.0793289047645905E-5, 1.0463173212266783E-5, 1.0139232120183559E-5, 9.8214558185907186E-6, 9.5098297263323067E-6, 9.20433485322091E-6, 8.9049480131616991E-6, 0.0, 0.0, 0.0, 0.0, -0.0, -0.0, -0.0, -0.0, -0.0, -0.0, -0.0, -0.0, -0.0, -0.0, -0.0, -0.0, -0.0, -0.0, -0.0, -0.0, -0.0, -0.0, -0.0, -0.0, -0.0, -0.0, -0.0, -0.0, -0.0, -0.0, -0.0, -0.0, -0.0, -0.0, -0.0, -0.0, -0.0, -0.0, -0.0, -0.0, -0.0, -0.0, -0.0, -0.0, -0.0, -0.0, -0.0, -0.0, -0.0, -0.0, -0.0, -0.0, -0.0, -0.0, -0.0, -0.0, -0.0, -0.0, -0.0, -0.0, -0.0, -0.0, -0.0, -0.0, -0.0, -0.0, -0.0, -0.0, -0.0, -0.0, -0.0, -0.0, -0.0, -0.0, -0.0, -0.0, -0.0, -0.0, -0.0, -0.0, -0.0, -0.0, -0.0, -0.0, -0.0, -0.0, -0.0, -0.0, -0.0, -0.0, -0.0, -0.0, -0.0, -0.0, -0.0, -0.0, -0.0, -0.0, -0.0, -0.0, -0.0, -0.0, -0.0, -0.0, -0.0, -0.0, -0.0, -0.0, -0.0, -0.0, -0.0, -0.0, -0.0, -0.0, -0.0, -0.0, -0.0, -0.0, -0.0, -0.0, -0.0, -0.0, -0.0, -0.0, 0.0, 0.0, 0.0, 0.0, 0.0, 0.0, 0.0, 0.0, 0.0, 0.0, 0.0, 0.0, 0.0, 0.0, 0.0, 0.0, 0.0, 0.0, 0.0, 0.0, 0.0, 0.0, 0.0, 0.0, 0.0, 0.0, 0.0, 0.0, 0.0, 0.0, 0.0, 0.0, 0.0, 0.0, 0.0, 0.0, 0.0, 0.0, 0.0, 0.0, 0.0, 0.0, 0.0, 0.0, 0.0, 0.0, 0.0, 0.0, 0.0, 0.0, 0.0, 0.0, 0.0, 0.0, 0.0, 0.0, 0.0, 0.0, 0.0, 0.0, 0.0, 0.0, 0.0, 0.0, 0.0, 0.0, 0.0, 0.0, 0.0, 0.0, 0.0, 0.0, 0.0, 0.0, 0.0, 0.0, 0.0, 0.0, 0.0, 0.0, 0.0, 0.0, 0.0, 0.0, 0.0, 0.0, 0.0, 0.0, 0.0, 0.0, 0.0, 0.0, 0.0, 0.0, 0.0, 0.0, 0.0, 0.0, 0.0, 0.0, 0.0, 0.0, 0.0, 0.0, 0.0, 0.0, 0.0, 0.0, 0.0, 0.0, 0.0, 0.0, 0.0, 0.0, 0.0, 0.0, 0.0, 0.0, 0.0, 0.0, 0.0, 0.0, 0.0, 0.0, -0.0, -0.0, -0.0, -0.0, -0.0, -0.0, -0.0, -0.0, -0.0, -0.0, -1.7756006070928429E-5, -1.955926027849794E-5, -2.1265642444599059E-5, -2.2878087249309936E-5, -2.4399475238503513E-5, -2.5832632877734329E-5, -2.7180332648224444E-5, -2.8445293182983732E-5, -2.9630179441154765E-5, -3.0737602918726609E-5, -3.1770121893815045E-5, -3.2730241704758869E-5, -3.3620415059333691E-5, -3.4443042373434618E-5, -3.5200472137629193E-5, -3.5895001310030509E-5, -3.652887573398812E-5, -3.7104290579141277E-5, -3.7623390804425058E-5, -3.808827164166491E-5, -3.8500979098439383E-5, -3.886351047893401E-5, -3.9177814921551905E-5, -3.9445793952087749E-5, -3.966930205131298E-5, -3.98501472358593E-5, -3.9990091651326829E-5, -4.0090852176581095E-5, -4.0154101038240283E-5, -4.0181466434390562E-5, -4.017453316660271E-5, -4.013484327935801E-5, -4.0063896706025282E-5, -3.9963151920563813E-5, -3.9834026594159355E-5, -3.9677898256031791E-5, -3.9496104957683613E-5, -3.9289945939888413E-5, -3.9060682301747689E-5, -3.8809537671172525E-5, -3.8537698876174604E-5, -3.8246316616377579E-5, -3.793650613418646E-5, -3.7609347885077623E-5, -3.7265888206497395E-5, -3.6907139984880808E-5, -3.6534083320325723E-5, -3.6147666188480321E-5, -3.5748805099224027E-5, -3.5338385751743129E-5, -3.4917263685623729E-5, -3.44862649276042E-5, -3.40461866336495E-5, -3.3597797726028135E-5, -3.3141839525091535E-5, -3.2679026375472935E-5, -3.221004626644033E-5, -3.1735561446154833E-5, -3.12562090296018E-5, -3.0772601599977736E-5, -3.0285327803331116E-5, -2.9794952936269942E-5, -2.9302019526562752E-5, -2.8807047906473585E-5, -2.8310536778684464E-5, -2.7812963774671571E-5, -2.7314786005413577E-5, -2.6816440604322343E-5, -2.6318345262297408E-5, -2.5820898754816765E-5, -2.5324481460986734E-5, -2.4829455874483883E-5, -2.4336167106331684E-5, -2.3844943379463754E-5, -2.3356096515034559E-5, -2.2869922410446928E-5, -2.2386701509073987E-5, -2.190669926166088E-5, -2.1430166579399207E-5, -2.0957340278674263E-5, -2.0488443517492027E-5, -2.0023686223599328E-5, -1.9563265514316956E-5, -1.910736610811127E-5, -1.8656160727935741E-5, -1.8209810496378919E-5, -1.776846532266075E-5, -1.7332264281523728E-5, -1.6901335984070202E-5, -1.6475798940601218E-5, -1.6055761915516631E-5, -1.5641324274339943E-5, -1.5232576322934952E-5, -1.4829599638984815E-5, -1.4432467395807249E-5, -1.4041244678582621E-5, -1.3655988793074526E-5, -1.3276749566924981E-5, -1.29035696436089E-5, -1.2536484769134677E-5, -1.217552407157984E-5, -1.1820710333552607E-5, -1.1472060257671982E-5, -1.1129584725160594E-5, -1.0793289047645905E-5, -1.0463173212266783E-5, -1.0139232120183559E-5, -9.8214558185907186E-6, -9.5098297263323067E-6, -9.20433485322091E-6, 0.0, 0.0, 0.0, 0.0, 0.0, 0.0, 0.0, 0.0, 0.0, 0.0, 1.7756006070928429E-5, 1.955926027849794E-5, 2.1265642444599059E-5, 2.2878087249309936E-5, 2.4399475238503513E-5, 2.5832632877734329E-5, 2.7180332648224444E-5, 2.8445293182983732E-5, 2.9630179441154765E-5, 3.0737602918726609E-5, 3.1770121893815045E-5, 3.2730241704758869E-5, 3.3620415059333691E-5, 3.4443042373434618E-5, 3.5200472137629193E-5, 3.5895001310030509E-5, 3.652887573398812E-5, 3.7104290579141277E-5, 3.7623390804425058E-5, 3.808827164166491E-5, 3.8500979098439383E-5, 3.886351047893401E-5, 3.9177814921551905E-5, 3.9445793952087749E-5, 3.966930205131298E-5, 3.98501472358593E-5, 3.9990091651326829E-5, 4.0090852176581095E-5, 4.0154101038240283E-5, 4.0181466434390562E-5, 4.017453316660271E-5, 4.013484327935801E-5, 4.0063896706025282E-5, 3.9963151920563813E-5, 3.9834026594159355E-5, 3.9677898256031791E-5, 3.9496104957683613E-5, 3.9289945939888413E-5, 3.9060682301747689E-5, 3.8809537671172525E-5, 3.8537698876174604E-5, 3.8246316616377579E-5, 3.793650613418646E-5, 3.7609347885077623E-5, 3.7265888206497395E-5, 3.6907139984880808E-5, 3.6534083320325723E-5, 3.6147666188480321E-5, 3.5748805099224027E-5, 3.5338385751743129E-5, 3.4917263685623729E-5, 3.44862649276042E-5, 3.40461866336495E-5, 3.3597797726028135E-5, 3.3141839525091535E-5, 3.2679026375472935E-5, 3.221004626644033E-5, 3.1735561446154833E-5, 3.12562090296018E-5, 3.0772601599977736E-5, 3.0285327803331116E-5, 2.9794952936269942E-5, 2.9302019526562752E-5, 2.8807047906473585E-5, 2.8310536778684464E-5, 2.7812963774671571E-5, 2.7314786005413577E-5, 2.6816440604322343E-5, 2.6318345262297408E-5, 2.5820898754816765E-5, 2.5324481460986734E-5, 2.4829455874483883E-5, 2.4336167106331684E-5, 2.3844943379463754E-5, 2.3356096515034559E-5, 2.2869922410446928E-5, 2.2386701509073987E-5, 2.190669926166088E-5, 2.1430166579399207E-5, 2.0957340278674263E-5, 2.0488443517492027E-5, 2.0023686223599328E-5, 1.9563265514316956E-5, 1.910736610811127E-5, 1.8656160727935741E-5, 1.8209810496378919E-5, 1.776846532266075E-5, 1.7332264281523728E-5, 1.6901335984070202E-5, 1.6475798940601218E-5, 1.6055761915516631E-5, 1.5641324274339943E-5, 1.5232576322934952E-5, 1.4829599638984815E-5, 1.4432467395807249E-5, 1.4041244678582621E-5, 1.3655988793074526E-5, 1.3276749566924981E-5, 1.29035696436089E-5, 1.2536484769134677E-5, 1.217552407157984E-5, 1.1820710333552607E-5, 1.1472060257671982E-5, 1.1129584725160594E-5, 1.0793289047645905E-5, 1.0463173212266783E-5, 1.0139232120183559E-5, 9.8214558185907186E-6, 9.5098297263323067E-6, 9.20433485322091E-6, 0.0, 0.0, 0.0, 0.0, -0.0, -0.0, -0.0, -0.0, -0.0, -0.0, -0.0, -0.0, -0.0, -0.0, -0.0, -0.0, -0.0, -0.0, -0.0, -0.0, -0.0, -0.0, -0.0, -0.0, -0.0, -0.0, -0.0, -0.0, -0.0, -0.0, -0.0, -0.0, -0.0, -0.0, -0.0, -0.0, -0.0, -0.0, -0.0, -0.0, -0.0, -0.0, -0.0, -0.0, -0.0, -0.0, -0.0, -0.0, -0.0, -0.0, -0.0, -0.0, -0.0, -0.0, -0.0, -0.0, -0.0, -0.0, -0.0, -0.0, -0.0, -0.0, -0.0, -0.0, -0.0, -0.0, -0.0, -0.0, -0.0, -0.0, -0.0, -0.0, -0.0, -0.0, -0.0, -0.0, -0.0, -0.0, -0.0, -0.0, -0.0, -0.0, -0.0, -0.0, -0.0, -0.0, -0.0, -0.0, -0.0, -0.0, -0.0, -0.0, -0.0, -0.0, -0.0, -0.0, -0.0, -0.0, -0.0, -0.0, -0.0, -0.0, -0.0, -0.0, -0.0, -0.0, -0.0, -0.0, -0.0, -0.0, -0.0, -0.0, -0.0, -0.0, -0.0, -0.0, -0.0, -0.0, -0.0, -0.0, -0.0, -0.0, -0.0, -0.0, 0.0, 0.0, 0.0, 0.0, 0.0, 0.0, 0.0, 0.0, 0.0, 0.0, 0.0, 0.0, 0.0, 0.0, 0.0, 0.0, 0.0, 0.0, 0.0, 0.0, 0.0, 0.0, 0.0, 0.0, 0.0, 0.0, 0.0, 0.0, 0.0, 0.0, 0.0, 0.0, 0.0, 0.0, 0.0, 0.0, 0.0, 0.0, 0.0, 0.0, 0.0, 0.0, 0.0, 0.0, 0.0, 0.0, 0.0, 0.0, 0.0, 0.0, 0.0, 0.0, 0.0, 0.0, 0.0, 0.0, 0.0, 0.0, 0.0, 0.0, 0.0, 0.0, 0.0, 0.0, 0.0, 0.0, 0.0, 0.0, 0.0, 0.0, 0.0, 0.0, 0.0, 0.0, 0.0, 0.0, 0.0, 0.0, 0.0, 0.0, 0.0, 0.0, 0.0, 0.0, 0.0, 0.0, 0.0, 0.0, 0.0, 0.0, 0.0, 0.0, 0.0, 0.0, 0.0, 0.0, 0.0, 0.0, 0.0, 0.0, 0.0, 0.0, 0.0, 0.0, 0.0, 0.0, 0.0, 0.0, 0.0, 0.0, 0.0, 0.0, 0.0, 0.0, 0.0, 0.0, 0.0, 0.0, 0.0, 0.0, 0.0, 0.0, 0.0, 0.0, -0.0, -0.0, -0.0, -0.0, -0.0, -0.0, -0.0, -0.0, -0.0, -0.0, -0.0, -1.7756006070928429E-5, -1.955926027849794E-5, -2.1265642444599059E-5, -2.2878087249309936E-5, -2.4399475238503513E-5, -2.5832632877734329E-5, -2.7180332648224444E-5, -2.8445293182983732E-5, -2.9630179441154765E-5, -3.0737602918726609E-5, -3.1770121893815045E-5, -3.2730241704758869E-5, -3.3620415059333691E-5, -3.4443042373434618E-5, -3.5200472137629193E-5, -3.5895001310030509E-5, -3.652887573398812E-5, -3.7104290579141277E-5, -3.7623390804425058E-5, -3.808827164166491E-5, -3.8500979098439383E-5, -3.886351047893401E-5, -3.9177814921551905E-5, -3.9445793952087749E-5, -3.966930205131298E-5, -3.98501472358593E-5, -3.9990091651326829E-5, -4.0090852176581095E-5, -4.0154101038240283E-5, -4.0181466434390562E-5, -4.017453316660271E-5, -4.013484327935801E-5, -4.0063896706025282E-5, -3.9963151920563813E-5, -3.9834026594159355E-5, -3.9677898256031791E-5, -3.9496104957683613E-5, -3.9289945939888413E-5, -3.9060682301747689E-5, -3.8809537671172525E-5, -3.8537698876174604E-5, -3.8246316616377579E-5, -3.793650613418646E-5, -3.7609347885077623E-5, -3.7265888206497395E-5, -3.6907139984880808E-5, -3.6534083320325723E-5, -3.6147666188480321E-5, -3.5748805099224027E-5, -3.5338385751743129E-5, -3.4917263685623729E-5, -3.44862649276042E-5, -3.40461866336495E-5, -3.3597797726028135E-5, -3.3141839525091535E-5, -3.2679026375472935E-5, -3.221004626644033E-5, -3.1735561446154833E-5, -3.12562090296018E-5, -3.0772601599977736E-5, -3.0285327803331116E-5, -2.9794952936269942E-5, -2.9302019526562752E-5, -2.8807047906473585E-5, -2.8310536778684464E-5, -2.7812963774671571E-5, -2.7314786005413577E-5, -2.6816440604322343E-5, -2.6318345262297408E-5, -2.5820898754816765E-5, -2.5324481460986734E-5, -2.4829455874483883E-5, -2.4336167106331684E-5, -2.3844943379463754E-5, -2.3356096515034559E-5, -2.2869922410446928E-5, -2.2386701509073987E-5, -2.190669926166088E-5, -2.1430166579399207E-5, -2.0957340278674263E-5, -2.0488443517492027E-5, -2.0023686223599328E-5, -1.9563265514316956E-5, -1.910736610811127E-5, -1.8656160727935741E-5, -1.8209810496378919E-5, -1.776846532266075E-5, -1.7332264281523728E-5, -1.6901335984070202E-5, -1.6475798940601218E-5, -1.6055761915516631E-5, -1.5641324274339943E-5, -1.5232576322934952E-5, -1.4829599638984815E-5, -1.4432467395807249E-5, -1.4041244678582621E-5, -1.3655988793074526E-5, -1.3276749566924981E-5, -1.29035696436089E-5, -1.2536484769134677E-5, -1.217552407157984E-5, -1.1820710333552607E-5, -1.1472060257671982E-5, -1.1129584725160594E-5, -1.0793289047645905E-5, -1.0463173212266783E-5, -1.0139232120183559E-5, -9.8214558185907186E-6, -9.5098297263323067E-6, 0.0, 0.0, 0.0, 0.0, 0.0, 0.0, 0.0, 0.0, 0.0, 0.0, 0.0, 1.7756006070928429E-5, 1.955926027849794E-5, 2.1265642444599059E-5, 2.2878087249309936E-5, 2.4399475238503513E-5, 2.5832632877734329E-5, 2.7180332648224444E-5, 2.8445293182983732E-5, 2.9630179441154765E-5, 3.0737602918726609E-5, 3.1770121893815045E-5, 3.2730241704758869E-5, 3.3620415059333691E-5, 3.4443042373434618E-5, 3.5200472137629193E-5, 3.5895001310030509E-5, 3.652887573398812E-5, 3.7104290579141277E-5, 3.7623390804425058E-5, 3.808827164166491E-5, 3.8500979098439383E-5, 3.886351047893401E-5, 3.9177814921551905E-5, 3.9445793952087749E-5, 3.966930205131298E-5, 3.98501472358593E-5, 3.9990091651326829E-5, 4.0090852176581095E-5, 4.0154101038240283E-5, 4.0181466434390562E-5, 4.017453316660271E-5, 4.013484327935801E-5, 4.0063896706025282E-5, 3.9963151920563813E-5, 3.9834026594159355E-5, 3.9677898256031791E-5, 3.9496104957683613E-5, 3.9289945939888413E-5, 3.9060682301747689E-5, 3.8809537671172525E-5, 3.8537698876174604E-5, 3.8246316616377579E-5, 3.793650613418646E-5, 3.7609347885077623E-5, 3.7265888206497395E-5, 3.6907139984880808E-5, 3.6534083320325723E-5, 3.6147666188480321E-5, 3.5748805099224027E-5, 3.5338385751743129E-5, 3.4917263685623729E-5, 3.44862649276042E-5, 3.40461866336495E-5, 3.3597797726028135E-5, 3.3141839525091535E-5, 3.2679026375472935E-5, 3.221004626644033E-5, 3.1735561446154833E-5, 3.12562090296018E-5, 3.0772601599977736E-5, 3.0285327803331116E-5, 2.9794952936269942E-5, 2.9302019526562752E-5, 2.8807047906473585E-5, 2.8310536778684464E-5, 2.7812963774671571E-5, 2.7314786005413577E-5, 2.6816440604322343E-5, 2.6318345262297408E-5, 2.5820898754816765E-5, 2.5324481460986734E-5, 2.4829455874483883E-5, 2.4336167106331684E-5, 2.3844943379463754E-5, 2.3356096515034559E-5, 2.2869922410446928E-5, 2.2386701509073987E-5, 2.190669926166088E-5, 2.1430166579399207E-5, 2.0957340278674263E-5, 2.0488443517492027E-5, 2.0023686223599328E-5, 1.9563265514316956E-5, 1.910736610811127E-5, 1.8656160727935741E-5, 1.8209810496378919E-5, 1.776846532266075E-5, 1.7332264281523728E-5, 1.6901335984070202E-5, 1.6475798940601218E-5, 1.6055761915516631E-5, 1.5641324274339943E-5, 1.5232576322934952E-5, 1.4829599638984815E-5, 1.4432467395807249E-5, 1.4041244678582621E-5, 1.3655988793074526E-5, 1.3276749566924981E-5, 1.29035696436089E-5, 1.2536484769134677E-5, 1.217552407157984E-5, 1.1820710333552607E-5, 1.1472060257671982E-5, 1.1129584725160594E-5, 1.0793289047645905E-5, 1.0463173212266783E-5, 1.0139232120183559E-5, 9.8214558185907186E-6, 9.5098297263323067E-6, 0.0, 0.0, 0.0, 0.0, -0.0, -0.0, -0.0, -0.0, -0.0, -0.0, -0.0, -0.0, -0.0, -0.0, -0.0, -0.0, -0.0, -0.0, -0.0, -0.0, -0.0, -0.0, -0.0, -0.0, -0.0, -0.0, -0.0, -0.0, -0.0, -0.0, -0.0, -0.0, -0.0, -0.0, -0.0, -0.0, -0.0, -0.0, -0.0, -0.0, -0.0, -0.0, -0.0, -0.0, -0.0, -0.0, -0.0, -0.0, -0.0, -0.0, -0.0, -0.0, -0.0, -0.0, -0.0, -0.0, -0.0, -0.0, -0.0, -0.0, -0.0, -0.0, -0.0, -0.0, -0.0, -0.0, -0.0, -0.0, -0.0, -0.0, -0.0, -0.0, -0.0, -0.0, -0.0, -0.0, -0.0, -0.0, -0.0, -0.0, -0.0, -0.0, -0.0, -0.0, -0.0, -0.0, -0.0, -0.0, -0.0, -0.0, -0.0, -0.0, -0.0, -0.0, -0.0, -0.0, -0.0, -0.0, -0.0, -0.0, -0.0, -0.0, -0.0, -0.0, -0.0, -0.0, -0.0, -0.0, -0.0, -0.0, -0.0, -0.0, -0.0, -0.0, -0.0, -0.0, -0.0, -0.0, -0.0, -0.0, -0.0, -0.0, -0.0, -0.0, 0.0, 0.0, 0.0, 0.0, 0.0, 0.0, 0.0, 0.0, 0.0, 0.0, 0.0, 0.0, 0.0, 0.0, 0.0, 0.0, 0.0, 0.0, 0.0, 0.0, 0.0, 0.0, 0.0, 0.0, 0.0, 0.0, 0.0, 0.0, 0.0, 0.0, 0.0, 0.0, 0.0, 0.0, 0.0, 0.0, 0.0, 0.0, 0.0, 0.0, 0.0, 0.0, 0.0, 0.0, 0.0, 0.0, 0.0, 0.0, 0.0, 0.0, 0.0, 0.0, 0.0, 0.0, 0.0, 0.0, 0.0, 0.0, 0.0, 0.0, 0.0, 0.0, 0.0, 0.0, 0.0, 0.0, 0.0, 0.0, 0.0, 0.0, 0.0, 0.0, 0.0, 0.0, 0.0, 0.0, 0.0, 0.0, 0.0, 0.0, 0.0, 0.0, 0.0, 0.0, 0.0, 0.0, 0.0, 0.0, 0.0, 0.0, 0.0, 0.0, 0.0, 0.0, 0.0, 0.0, 0.0, 0.0, 0.0, 0.0, 0.0, 0.0, 0.0, 0.0, 0.0, 0.0, 0.0, 0.0, 0.0, 0.0, 0.0, 0.0, 0.0, 0.0, 0.0, 0.0, 0.0, 0.0, 0.0, 0.0, 0.0, 0.0, 0.0, 0.0, -0.0, -0.0, -0.0, -0.0, -0.0, -0.0, -0.0, -0.0, -0.0, -0.0, -0.0, -0.0, -1.7756006070928429E-5, -1.955926027849794E-5, -2.1265642444599059E-5, -2.2878087249309936E-5, -2.4399475238503513E-5, -2.5832632877734329E-5, -2.7180332648224444E-5, -2.8445293182983732E-5, -2.9630179441154765E-5, -3.0737602918726609E-5, -3.1770121893815045E-5, -3.2730241704758869E-5, -3.3620415059333691E-5, -3.4443042373434618E-5, -3.5200472137629193E-5, -3.5895001310030509E-5, -3.652887573398812E-5, -3.7104290579141277E-5, -3.7623390804425058E-5, -3.808827164166491E-5, -3.8500979098439383E-5, -3.886351047893401E-5, -3.9177814921551905E-5, -3.9445793952087749E-5, -3.966930205131298E-5, -3.98501472358593E-5, -3.9990091651326829E-5, -4.0090852176581095E-5, -4.0154101038240283E-5, -4.0181466434390562E-5, -4.017453316660271E-5, -4.013484327935801E-5, -4.0063896706025282E-5, -3.9963151920563813E-5, -3.9834026594159355E-5, -3.9677898256031791E-5, -3.9496104957683613E-5, -3.9289945939888413E-5, -3.9060682301747689E-5, -3.8809537671172525E-5, -3.8537698876174604E-5, -3.8246316616377579E-5, -3.793650613418646E-5, -3.7609347885077623E-5, -3.7265888206497395E-5, -3.6907139984880808E-5, -3.6534083320325723E-5, -3.6147666188480321E-5, -3.5748805099224027E-5, -3.5338385751743129E-5, -3.4917263685623729E-5, -3.44862649276042E-5, -3.40461866336495E-5, -3.3597797726028135E-5, -3.3141839525091535E-5, -3.2679026375472935E-5, -3.221004626644033E-5, -3.1735561446154833E-5, -3.12562090296018E-5, -3.0772601599977736E-5, -3.0285327803331116E-5, -2.9794952936269942E-5, -2.9302019526562752E-5, -2.8807047906473585E-5, -2.8310536778684464E-5, -2.7812963774671571E-5, -2.7314786005413577E-5, -2.6816440604322343E-5, -2.6318345262297408E-5, -2.5820898754816765E-5, -2.5324481460986734E-5, -2.4829455874483883E-5, -2.4336167106331684E-5, -2.3844943379463754E-5, -2.3356096515034559E-5, -2.2869922410446928E-5, -2.2386701509073987E-5, -2.190669926166088E-5, -2.1430166579399207E-5, -2.0957340278674263E-5, -2.0488443517492027E-5, -2.0023686223599328E-5, -1.9563265514316956E-5, -1.910736610811127E-5, -1.8656160727935741E-5, -1.8209810496378919E-5, -1.776846532266075E-5, -1.7332264281523728E-5, -1.6901335984070202E-5, -1.6475798940601218E-5, -1.6055761915516631E-5, -1.5641324274339943E-5, -1.5232576322934952E-5, -1.4829599638984815E-5, -1.4432467395807249E-5, -1.4041244678582621E-5, -1.3655988793074526E-5, -1.3276749566924981E-5, -1.29035696436089E-5, -1.2536484769134677E-5, -1.217552407157984E-5, -1.1820710333552607E-5, -1.1472060257671982E-5, -1.1129584725160594E-5, -1.0793289047645905E-5, -1.0463173212266783E-5, -1.0139232120183559E-5, -9.8214558185907186E-6, 0.0, 0.0, 0.0, 0.0, 0.0, 0.0, 0.0, 0.0, 0.0, 0.0, 0.0, 0.0, 1.7756006070928429E-5, 1.955926027849794E-5, 2.1265642444599059E-5, 2.2878087249309936E-5, 2.4399475238503513E-5, 2.5832632877734329E-5, 2.7180332648224444E-5, 2.8445293182983732E-5, 2.9630179441154765E-5, 3.0737602918726609E-5, 3.1770121893815045E-5, 3.2730241704758869E-5, 3.3620415059333691E-5, 3.4443042373434618E-5, 3.5200472137629193E-5, 3.5895001310030509E-5, 3.652887573398812E-5, 3.7104290579141277E-5, 3.7623390804425058E-5, 3.808827164166491E-5, 3.8500979098439383E-5, 3.886351047893401E-5, 3.9177814921551905E-5, 3.9445793952087749E-5, 3.966930205131298E-5, 3.98501472358593E-5, 3.9990091651326829E-5, 4.0090852176581095E-5, 4.0154101038240283E-5, 4.0181466434390562E-5, 4.017453316660271E-5, 4.013484327935801E-5, 4.0063896706025282E-5, 3.9963151920563813E-5, 3.9834026594159355E-5, 3.9677898256031791E-5, 3.9496104957683613E-5, 3.9289945939888413E-5, 3.9060682301747689E-5, 3.8809537671172525E-5, 3.8537698876174604E-5, 3.8246316616377579E-5, 3.793650613418646E-5, 3.7609347885077623E-5, 3.7265888206497395E-5, 3.6907139984880808E-5, 3.6534083320325723E-5, 3.6147666188480321E-5, 3.5748805099224027E-5, 3.5338385751743129E-5, 3.4917263685623729E-5, 3.44862649276042E-5, 3.40461866336495E-5, 3.3597797726028135E-5, 3.3141839525091535E-5, 3.2679026375472935E-5, 3.221004626644033E-5, 3.1735561446154833E-5, 3.12562090296018E-5, 3.0772601599977736E-5, 3.0285327803331116E-5, 2.9794952936269942E-5, 2.9302019526562752E-5, 2.8807047906473585E-5, 2.8310536778684464E-5, 2.7812963774671571E-5, 2.7314786005413577E-5, 2.6816440604322343E-5, 2.6318345262297408E-5, 2.5820898754816765E-5, 2.5324481460986734E-5, 2.4829455874483883E-5, 2.4336167106331684E-5, 2.3844943379463754E-5, 2.3356096515034559E-5, 2.2869922410446928E-5, 2.2386701509073987E-5, 2.190669926166088E-5, 2.1430166579399207E-5, 2.0957340278674263E-5, 2.0488443517492027E-5, 2.0023686223599328E-5, 1.9563265514316956E-5, 1.910736610811127E-5, 1.8656160727935741E-5, 1.8209810496378919E-5, 1.776846532266075E-5, 1.7332264281523728E-5, 1.6901335984070202E-5, 1.6475798940601218E-5, 1.6055761915516631E-5, 1.5641324274339943E-5, 1.5232576322934952E-5, 1.4829599638984815E-5, 1.4432467395807249E-5, 1.4041244678582621E-5, 1.3655988793074526E-5, 1.3276749566924981E-5, 1.29035696436089E-5, 1.2536484769134677E-5, 1.217552407157984E-5, 1.1820710333552607E-5, 1.1472060257671982E-5, 1.1129584725160594E-5, 1.0793289047645905E-5, 1.0463173212266783E-5, 1.0139232120183559E-5, 9.8214558185907186E-6, 0.0, 0.0, 0.0, 0.0, -0.0, -0.0, -0.0, -0.0, -0.0, -0.0, -0.0, -0.0, -0.0, -0.0, -0.0, -0.0, -0.0, -0.0, -0.0, -0.0, -0.0, -0.0, -0.0, -0.0, -0.0, -0.0, -0.0, -0.0, -0.0, -0.0, -0.0, -0.0, -0.0, -0.0, -0.0, -0.0, -0.0, -0.0, -0.0, -0.0, -0.0, -0.0, -0.0, -0.0, -0.0, -0.0, -0.0, -0.0, -0.0, -0.0, -0.0, -0.0, -0.0, -0.0, -0.0, -0.0, -0.0, -0.0, -0.0, -0.0, -0.0, -0.0, -0.0, -0.0, -0.0, -0.0, -0.0, -0.0, -0.0, -0.0, -0.0, -0.0, -0.0, -0.0, -0.0, -0.0, -0.0, -0.0, -0.0, -0.0, -0.0, -0.0, -0.0, -0.0, -0.0, -0.0, -0.0, -0.0, -0.0, -0.0, -0.0, -0.0, -0.0, -0.0, -0.0, -0.0, -0.0, -0.0, -0.0, -0.0, -0.0, -0.0, -0.0, -0.0, -0.0, -0.0, -0.0, -0.0, -0.0, -0.0, -0.0, -0.0, -0.0, -0.0, -0.0, -0.0, -0.0, -0.0, -0.0, -0.0, -0.0, -0.0, -0.0, -0.0, 0.0, 0.0, 0.0, 0.0, 0.0, 0.0, 0.0, 0.0, 0.0, 0.0, 0.0, 0.0, 0.0, 0.0, 0.0, 0.0, 0.0, 0.0, 0.0, 0.0, 0.0, 0.0, 0.0, 0.0, 0.0, 0.0, 0.0, 0.0, 0.0, 0.0, 0.0, 0.0, 0.0, 0.0, 0.0, 0.0, 0.0, 0.0, 0.0, 0.0, 0.0, 0.0, 0.0, 0.0, 0.0, 0.0, 0.0, 0.0, 0.0, 0.0, 0.0, 0.0, 0.0, 0.0, 0.0, 0.0, 0.0, 0.0, 0.0, 0.0, 0.0, 0.0, 0.0, 0.0, 0.0, 0.0, 0.0, 0.0, 0.0, 0.0, 0.0, 0.0, 0.0, 0.0, 0.0, 0.0, 0.0, 0.0, 0.0, 0.0, 0.0, 0.0, 0.0, 0.0, 0.0, 0.0, 0.0, 0.0, 0.0, 0.0, 0.0, 0.0, 0.0, 0.0, 0.0, 0.0, 0.0, 0.0, 0.0, 0.0, 0.0, 0.0, 0.0, 0.0, 0.0, 0.0, 0.0, 0.0, 0.0, 0.0, 0.0, 0.0, 0.0, 0.0, 0.0, 0.0, 0.0, 0.0, 0.0, 0.0, 0.0, 0.0, 0.0, 0.0, -0.0, -0.0, -0.0, -0.0, -0.0, -0.0, -0.0, -0.0, -0.0, -0.0, -0.0, -0.0, -0.0, -1.7756006070928429E-5, -1.955926027849794E-5, -2.1265642444599059E-5, -2.2878087249309936E-5, -2.4399475238503513E-5, -2.5832632877734329E-5, -2.7180332648224444E-5, -2.8445293182983732E-5, -2.9630179441154765E-5, -3.0737602918726609E-5, -3.1770121893815045E-5, -3.2730241704758869E-5, -3.3620415059333691E-5, -3.4443042373434618E-5, -3.5200472137629193E-5, -3.5895001310030509E-5, -3.652887573398812E-5, -3.7104290579141277E-5, -3.7623390804425058E-5, -3.808827164166491E-5, -3.8500979098439383E-5, -3.886351047893401E-5, -3.9177814921551905E-5, -3.9445793952087749E-5, -3.966930205131298E-5, -3.98501472358593E-5, -3.9990091651326829E-5, -4.0090852176581095E-5, -4.0154101038240283E-5, -4.0181466434390562E-5, -4.017453316660271E-5, -4.013484327935801E-5, -4.0063896706025282E-5, -3.9963151920563813E-5, -3.9834026594159355E-5, -3.9677898256031791E-5, -3.9496104957683613E-5, -3.9289945939888413E-5, -3.9060682301747689E-5, -3.8809537671172525E-5, -3.8537698876174604E-5, -3.8246316616377579E-5, -3.793650613418646E-5, -3.7609347885077623E-5, -3.7265888206497395E-5, -3.6907139984880808E-5, -3.6534083320325723E-5, -3.6147666188480321E-5, -3.5748805099224027E-5, -3.5338385751743129E-5, -3.4917263685623729E-5, -3.44862649276042E-5, -3.40461866336495E-5, -3.3597797726028135E-5, -3.3141839525091535E-5, -3.2679026375472935E-5, -3.221004626644033E-5, -3.1735561446154833E-5, -3.12562090296018E-5, -3.0772601599977736E-5, -3.0285327803331116E-5, -2.9794952936269942E-5, -2.9302019526562752E-5, -2.8807047906473585E-5, -2.8310536778684464E-5, -2.7812963774671571E-5, -2.7314786005413577E-5, -2.6816440604322343E-5, -2.6318345262297408E-5, -2.5820898754816765E-5, -2.5324481460986734E-5, -2.4829455874483883E-5, -2.4336167106331684E-5, -2.3844943379463754E-5, -2.3356096515034559E-5, -2.2869922410446928E-5, -2.2386701509073987E-5, -2.190669926166088E-5, -2.1430166579399207E-5, -2.0957340278674263E-5, -2.0488443517492027E-5, -2.0023686223599328E-5, -1.9563265514316956E-5, -1.910736610811127E-5, -1.8656160727935741E-5, -1.8209810496378919E-5, -1.776846532266075E-5, -1.7332264281523728E-5, -1.6901335984070202E-5, -1.6475798940601218E-5, -1.6055761915516631E-5, -1.5641324274339943E-5, -1.5232576322934952E-5, -1.4829599638984815E-5, -1.4432467395807249E-5, -1.4041244678582621E-5, -1.3655988793074526E-5, -1.3276749566924981E-5, -1.29035696436089E-5, -1.2536484769134677E-5, -1.217552407157984E-5, -1.1820710333552607E-5, -1.1472060257671982E-5, -1.1129584725160594E-5, -1.0793289047645905E-5, -1.0463173212266783E-5, -1.0139232120183559E-5, 0.0, 0.0, 0.0, 0.0, 0.0, 0.0, 0.0, 0.0, 0.0, 0.0, 0.0, 0.0, 0.0, 1.7756006070928429E-5, 1.955926027849794E-5, 2.1265642444599059E-5, 2.2878087249309936E-5, 2.4399475238503513E-5, 2.5832632877734329E-5, 2.7180332648224444E-5, 2.8445293182983732E-5, 2.9630179441154765E-5, 3.0737602918726609E-5, 3.1770121893815045E-5, 3.2730241704758869E-5, 3.3620415059333691E-5, 3.4443042373434618E-5, 3.5200472137629193E-5, 3.5895001310030509E-5, 3.652887573398812E-5, 3.7104290579141277E-5, 3.7623390804425058E-5, 3.808827164166491E-5, 3.8500979098439383E-5, 3.886351047893401E-5, 3.9177814921551905E-5, 3.9445793952087749E-5, 3.966930205131298E-5, 3.98501472358593E-5, 3.9990091651326829E-5, 4.0090852176581095E-5, 4.0154101038240283E-5, 4.0181466434390562E-5, 4.017453316660271E-5, 4.013484327935801E-5, 4.0063896706025282E-5, 3.9963151920563813E-5, 3.9834026594159355E-5, 3.9677898256031791E-5, 3.9496104957683613E-5, 3.9289945939888413E-5, 3.9060682301747689E-5, 3.8809537671172525E-5, 3.8537698876174604E-5, 3.8246316616377579E-5, 3.793650613418646E-5, 3.7609347885077623E-5, 3.7265888206497395E-5, 3.6907139984880808E-5, 3.6534083320325723E-5, 3.6147666188480321E-5, 3.5748805099224027E-5, 3.5338385751743129E-5, 3.4917263685623729E-5, 3.44862649276042E-5, 3.40461866336495E-5, 3.3597797726028135E-5, 3.3141839525091535E-5, 3.2679026375472935E-5, 3.221004626644033E-5, 3.1735561446154833E-5, 3.12562090296018E-5, 3.0772601599977736E-5, 3.0285327803331116E-5, 2.9794952936269942E-5, 2.9302019526562752E-5, 2.8807047906473585E-5, 2.8310536778684464E-5, 2.7812963774671571E-5, 2.7314786005413577E-5, 2.6816440604322343E-5, 2.6318345262297408E-5, 2.5820898754816765E-5, 2.5324481460986734E-5, 2.4829455874483883E-5, 2.4336167106331684E-5, 2.3844943379463754E-5, 2.3356096515034559E-5, 2.2869922410446928E-5, 2.2386701509073987E-5, 2.190669926166088E-5, 2.1430166579399207E-5, 2.0957340278674263E-5, 2.0488443517492027E-5, 2.0023686223599328E-5, 1.9563265514316956E-5, 1.910736610811127E-5, 1.8656160727935741E-5, 1.8209810496378919E-5, 1.776846532266075E-5, 1.7332264281523728E-5, 1.6901335984070202E-5, 1.6475798940601218E-5, 1.6055761915516631E-5, 1.5641324274339943E-5, 1.5232576322934952E-5, 1.4829599638984815E-5, 1.4432467395807249E-5, 1.4041244678582621E-5, 1.3655988793074526E-5, 1.3276749566924981E-5, 1.29035696436089E-5, 1.2536484769134677E-5, 1.217552407157984E-5, 1.1820710333552607E-5, 1.1472060257671982E-5, 1.1129584725160594E-5, 1.0793289047645905E-5, 1.0463173212266783E-5, 1.0139232120183559E-5, 0.0, 0.0, 0.0, 0.0, -0.0, -0.0, -0.0, -0.0, -0.0, -0.0, -0.0, -0.0, -0.0, -0.0, -0.0, -0.0, -0.0, -0.0, -0.0, -0.0, -0.0, -0.0, -0.0, -0.0, -0.0, -0.0, -0.0, -0.0, -0.0, -0.0, -0.0, -0.0, -0.0, -0.0, -0.0, -0.0, -0.0, -0.0, -0.0, -0.0, -0.0, -0.0, -0.0, -0.0, -0.0, -0.0, -0.0, -0.0, -0.0, -0.0, -0.0, -0.0, -0.0, -0.0, -0.0, -0.0, -0.0, -0.0, -0.0, -0.0, -0.0, -0.0, -0.0, -0.0, -0.0, -0.0, -0.0, -0.0, -0.0, -0.0, -0.0, -0.0, -0.0, -0.0, -0.0, -0.0, -0.0, -0.0, -0.0, -0.0, -0.0, -0.0, -0.0, -0.0, -0.0, -0.0, -0.0, -0.0, -0.0, -0.0, -0.0, -0.0, -0.0, -0.0, -0.0, -0.0, -0.0, -0.0, -0.0, -0.0, -0.0, -0.0, -0.0, -0.0, -0.0, -0.0, -0.0, -0.0, -0.0, -0.0, -0.0, -0.0, -0.0, -0.0, -0.0, -0.0, -0.0, -0.0, -0.0, -0.0, -0.0, -0.0, -0.0, -0.0, 0.0, 0.0, 0.0, 0.0, 0.0, 0.0, 0.0, 0.0, 0.0, 0.0, 0.0, 0.0, 0.0, 0.0, 0.0, 0.0, 0.0, 0.0, 0.0, 0.0, 0.0, 0.0, 0.0, 0.0, 0.0, 0.0, 0.0, 0.0, 0.0, 0.0, 0.0, 0.0, 0.0, 0.0, 0.0, 0.0, 0.0, 0.0, 0.0, 0.0, 0.0, 0.0, 0.0, 0.0, 0.0, 0.0, 0.0, 0.0, 0.0, 0.0, 0.0, 0.0, 0.0, 0.0, 0.0, 0.0, 0.0, 0.0, 0.0, 0.0, 0.0, 0.0, 0.0, 0.0, 0.0, 0.0, 0.0, 0.0, 0.0, 0.0, 0.0, 0.0, 0.0, 0.0, 0.0, 0.0, 0.0, 0.0, 0.0, 0.0, 0.0, 0.0, 0.0, 0.0, 0.0, 0.0, 0.0, 0.0, 0.0, 0.0, 0.0, 0.0, 0.0, 0.0, 0.0, 0.0, 0.0, 0.0, 0.0, 0.0, 0.0, 0.0, 0.0, 0.0, 0.0, 0.0, 0.0, 0.0, 0.0, 0.0, 0.0, 0.0, 0.0, 0.0, 0.0, 0.0, 0.0, 0.0, 0.0, 0.0, 0.0, 0.0, 0.0, 0.0, -0.0, -0.0, -0.0, -0.0, -0.0, -0.0, -0.0, -0.0, -0.0, -0.0, -0.0, -0.0, -0.0, -0.0, -1.7756006070928429E-5, -1.955926027849794E-5, -2.1265642444599059E-5, -2.2878087249309936E-5, -2.4399475238503513E-5, -2.5832632877734329E-5, -2.7180332648224444E-5, -2.8445293182983732E-5, -2.9630179441154765E-5, -3.0737602918726609E-5, -3.1770121893815045E-5, -3.2730241704758869E-5, -3.3620415059333691E-5, -3.4443042373434618E-5, -3.5200472137629193E-5, -3.5895001310030509E-5, -3.652887573398812E-5, -3.7104290579141277E-5, -3.7623390804425058E-5, -3.808827164166491E-5, -3.8500979098439383E-5, -3.886351047893401E-5, -3.9177814921551905E-5, -3.9445793952087749E-5, -3.966930205131298E-5, -3.98501472358593E-5, -3.9990091651326829E-5, -4.0090852176581095E-5, -4.0154101038240283E-5, -4.0181466434390562E-5, -4.017453316660271E-5, -4.013484327935801E-5, -4.0063896706025282E-5, -3.9963151920563813E-5, -3.9834026594159355E-5, -3.9677898256031791E-5, -3.9496104957683613E-5, -3.9289945939888413E-5, -3.9060682301747689E-5, -3.8809537671172525E-5, -3.8537698876174604E-5, -3.8246316616377579E-5, -3.793650613418646E-5, -3.7609347885077623E-5, -3.7265888206497395E-5, -3.6907139984880808E-5, -3.6534083320325723E-5, -3.6147666188480321E-5, -3.5748805099224027E-5, -3.5338385751743129E-5, -3.4917263685623729E-5, -3.44862649276042E-5, -3.40461866336495E-5, -3.3597797726028135E-5, -3.3141839525091535E-5, -3.2679026375472935E-5, -3.221004626644033E-5, -3.1735561446154833E-5, -3.12562090296018E-5, -3.0772601599977736E-5, -3.0285327803331116E-5, -2.9794952936269942E-5, -2.9302019526562752E-5, -2.8807047906473585E-5, -2.8310536778684464E-5, -2.7812963774671571E-5, -2.7314786005413577E-5, -2.6816440604322343E-5, -2.6318345262297408E-5, -2.5820898754816765E-5, -2.5324481460986734E-5, -2.4829455874483883E-5, -2.4336167106331684E-5, -2.3844943379463754E-5, -2.3356096515034559E-5, -2.2869922410446928E-5, -2.2386701509073987E-5, -2.190669926166088E-5, -2.1430166579399207E-5, -2.0957340278674263E-5, -2.0488443517492027E-5, -2.0023686223599328E-5, -1.9563265514316956E-5, -1.910736610811127E-5, -1.8656160727935741E-5, -1.8209810496378919E-5, -1.776846532266075E-5, -1.7332264281523728E-5, -1.6901335984070202E-5, -1.6475798940601218E-5, -1.6055761915516631E-5, -1.5641324274339943E-5, -1.5232576322934952E-5, -1.4829599638984815E-5, -1.4432467395807249E-5, -1.4041244678582621E-5, -1.3655988793074526E-5, -1.3276749566924981E-5, -1.29035696436089E-5, -1.2536484769134677E-5, -1.217552407157984E-5, -1.1820710333552607E-5, -1.1472060257671982E-5, -1.1129584725160594E-5, -1.0793289047645905E-5, -1.0463173212266783E-5, 0.0, 0.0, 0.0, 0.0, 0.0, 0.0, 0.0, 0.0, 0.0, 0.0, 0.0, 0.0, 0.0, 0.0, 1.7756006070928429E-5, 1.955926027849794E-5, 2.1265642444599059E-5, 2.2878087249309936E-5, 2.4399475238503513E-5, 2.5832632877734329E-5, 2.7180332648224444E-5, 2.8445293182983732E-5, 2.9630179441154765E-5, 3.0737602918726609E-5, 3.1770121893815045E-5, 3.2730241704758869E-5, 3.3620415059333691E-5, 3.4443042373434618E-5, 3.5200472137629193E-5, 3.5895001310030509E-5, 3.652887573398812E-5, 3.7104290579141277E-5, 3.7623390804425058E-5, 3.808827164166491E-5, 3.8500979098439383E-5, 3.886351047893401E-5, 3.9177814921551905E-5, 3.9445793952087749E-5, 3.966930205131298E-5, 3.98501472358593E-5, 3.9990091651326829E-5, 4.0090852176581095E-5, 4.0154101038240283E-5, 4.0181466434390562E-5, 4.017453316660271E-5, 4.013484327935801E-5, 4.0063896706025282E-5, 3.9963151920563813E-5, 3.9834026594159355E-5, 3.9677898256031791E-5, 3.9496104957683613E-5, 3.9289945939888413E-5, 3.9060682301747689E-5, 3.8809537671172525E-5, 3.8537698876174604E-5, 3.8246316616377579E-5, 3.793650613418646E-5, 3.7609347885077623E-5, 3.7265888206497395E-5, 3.6907139984880808E-5, 3.6534083320325723E-5, 3.6147666188480321E-5, 3.5748805099224027E-5, 3.5338385751743129E-5, 3.4917263685623729E-5, 3.44862649276042E-5, 3.40461866336495E-5, 3.3597797726028135E-5, 3.3141839525091535E-5, 3.2679026375472935E-5, 3.221004626644033E-5, 3.1735561446154833E-5, 3.12562090296018E-5, 3.0772601599977736E-5, 3.0285327803331116E-5, 2.9794952936269942E-5, 2.9302019526562752E-5, 2.8807047906473585E-5, 2.8310536778684464E-5, 2.7812963774671571E-5, 2.7314786005413577E-5, 2.6816440604322343E-5, 2.6318345262297408E-5, 2.5820898754816765E-5, 2.5324481460986734E-5, 2.4829455874483883E-5, 2.4336167106331684E-5, 2.3844943379463754E-5, 2.3356096515034559E-5, 2.2869922410446928E-5, 2.2386701509073987E-5, 2.190669926166088E-5, 2.1430166579399207E-5, 2.0957340278674263E-5, 2.0488443517492027E-5, 2.0023686223599328E-5, 1.9563265514316956E-5, 1.910736610811127E-5, 1.8656160727935741E-5, 1.8209810496378919E-5, 1.776846532266075E-5, 1.7332264281523728E-5, 1.6901335984070202E-5, 1.6475798940601218E-5, 1.6055761915516631E-5, 1.5641324274339943E-5, 1.5232576322934952E-5, 1.4829599638984815E-5, 1.4432467395807249E-5, 1.4041244678582621E-5, 1.3655988793074526E-5, 1.3276749566924981E-5, 1.29035696436089E-5, 1.2536484769134677E-5, 1.217552407157984E-5, 1.1820710333552607E-5, 1.1472060257671982E-5, 1.1129584725160594E-5, 1.0793289047645905E-5, 1.0463173212266783E-5, 0.0, 0.0, 0.0, 0.0, -0.0, -0.0, -0.0, -0.0, -0.0, -0.0, -0.0, -0.0, -0.0, -0.0, -0.0, -0.0, -0.0, -0.0, -0.0, -0.0, -0.0, -0.0, -0.0, -0.0, -0.0, -0.0, -0.0, -0.0, -0.0, -0.0, -0.0, -0.0, -0.0, -0.0, -0.0, -0.0, -0.0, -0.0, -0.0, -0.0, -0.0, -0.0, -0.0, -0.0, -0.0, -0.0, -0.0, -0.0, -0.0, -0.0, -0.0, -0.0, -0.0, -0.0, -0.0, -0.0, -0.0, -0.0, -0.0, -0.0, -0.0, -0.0, -0.0, -0.0, -0.0, -0.0, -0.0, -0.0, -0.0, -0.0, -0.0, -0.0, -0.0, -0.0, -0.0, -0.0, -0.0, -0.0, -0.0, -0.0, -0.0, -0.0, -0.0, -0.0, -0.0, -0.0, -0.0, -0.0, -0.0, -0.0, -0.0, -0.0, -0.0, -0.0, -0.0, -0.0, -0.0, -0.0, -0.0, -0.0, -0.0, -0.0, -0.0, -0.0, -0.0, -0.0, -0.0, -0.0, -0.0, -0.0, -0.0, -0.0, -0.0, -0.0, -0.0, -0.0, -0.0, -0.0, -0.0, -0.0, -0.0, -0.0, -0.0, -0.0, 0.0, 0.0, 0.0, 0.0, 0.0, 0.0, 0.0, 0.0, 0.0, 0.0, 0.0, 0.0, 0.0, 0.0, 0.0, 0.0, 0.0, 0.0, 0.0, 0.0, 0.0, 0.0, 0.0, 0.0, 0.0, 0.0, 0.0, 0.0, 